REGION Network 4: alarmy
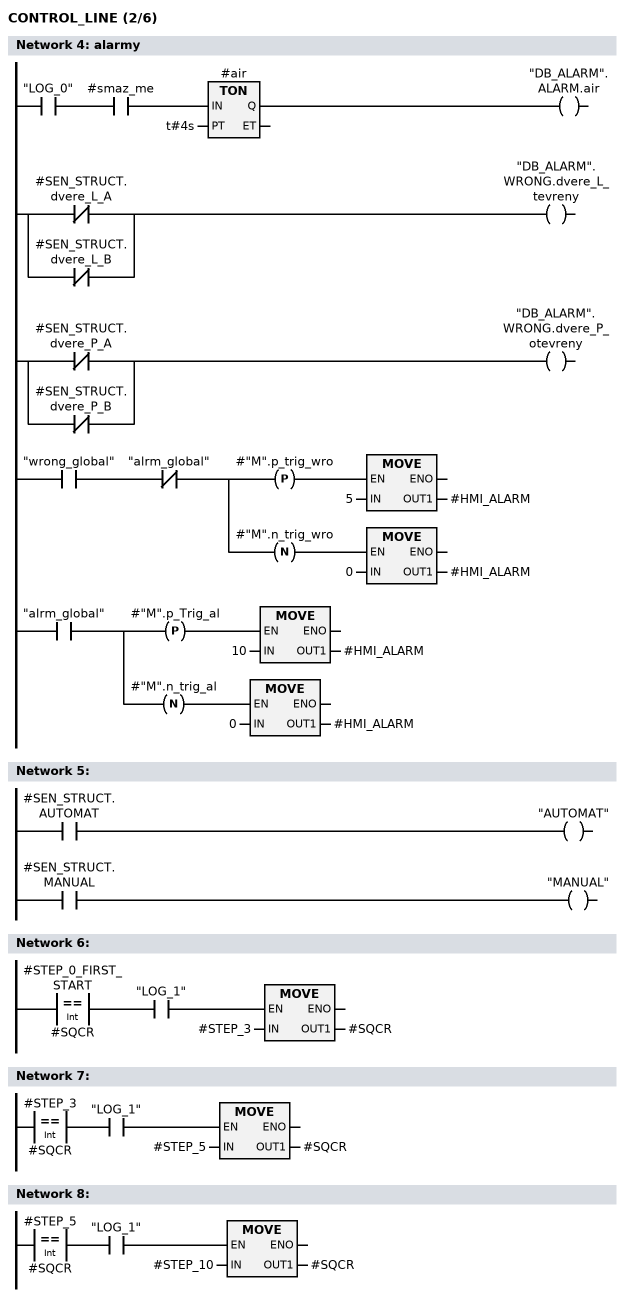
   #air(IN := "LOG_0" AND #smaz_me, PT := t#4s);   // TON
   "DB_ALARM".ALARM.air := #air.Q;
   "DB_ALARM".WRONG.dvere_L_tevreny := NOT #SEN_STRUCT.dvere_L_A OR NOT #SEN_STRUCT.dvere_L_B;
   "DB_ALARM".WRONG.dvere_P_otevreny := NOT #SEN_STRUCT.dvere_P_A OR NOT #SEN_STRUCT.dvere_P_B;
   #_w1 := "wrong_global" AND NOT "alrm_global";
   #_w2 := #_w1 AND NOT #"M".p_trig_wro;   // rising edge
   #"M".p_trig_wro := #_w1;
   IF #_w2 THEN #HMI_ALARM := 5; END_IF;
   #_w3 := NOT #_w1 AND #"M".n_trig_wro;   // falling edge
   #"M".n_trig_wro := #_w1;
   IF #_w3 THEN #HMI_ALARM := 0; END_IF;
   #_w4 := "alrm_global" AND NOT #"M".p_Trig_al;   // rising edge
   #"M".p_Trig_al := "alrm_global";
   IF #_w4 THEN #HMI_ALARM := 10; END_IF;
   #_w5 := NOT "alrm_global" AND #"M".n_trig_al;   // falling edge
   #"M".n_trig_al := "alrm_global";
   IF #_w5 THEN #HMI_ALARM := 0; END_IF;
END_REGION

REGION Network 5
   RUNG wire#powerrail
      Contact( #SEN_STRUCT.AUTOMAT )
      Coil( "AUTOMAT" )
   END_RUNG
   RUNG wire#powerrail
      Contact( #SEN_STRUCT.MANUAL )
      Coil( "MANUAL" )
   END_RUNG
   // the same network as SCL:
   "AUTOMAT" := #SEN_STRUCT.AUTOMAT;
   "MANUAL" := #SEN_STRUCT.MANUAL;
END_REGION

REGION Network 6
   RUNG wire#powerrail
      { S7_Templates := "SrcType := Int" } EQ_Contact(in1 := #STEP_0_FIRST_START, in2 := #SQCR)
      Contact( "LOG_1" )
      Move(in := #STEP_3, out1 => #SQCR)
   END_RUNG
   // the same network as SCL:
   IF (#STEP_0_FIRST_START = #SQCR) AND "LOG_1" THEN #SQCR := #STEP_3; END_IF;
END_REGION

REGION Network 7
   RUNG wire#powerrail
      { S7_Templates := "SrcType := Int" } EQ_Contact(in1 := #STEP_3, in2 := #SQCR)
      Contact( "LOG_1" )
      Move(in := #STEP_5, out1 => #SQCR)
   END_RUNG
   // the same network as SCL:
   IF (#STEP_3 = #SQCR) AND "LOG_1" THEN #SQCR := #STEP_5; END_IF;
END_REGION

REGION Network 8
   RUNG wire#powerrail
      { S7_Templates := "SrcType := Int" } EQ_Contact(in1 := #STEP_5, in2 := #SQCR)
      Contact( "LOG_1" )
      Move(in := #STEP_10, out1 => #SQCR)
   END_RUNG
   // the same network as SCL:
   IF (#STEP_5 = #SQCR) AND "LOG_1" THEN #SQCR := #STEP_10; END_IF;
END_REGION

REGION Network 9
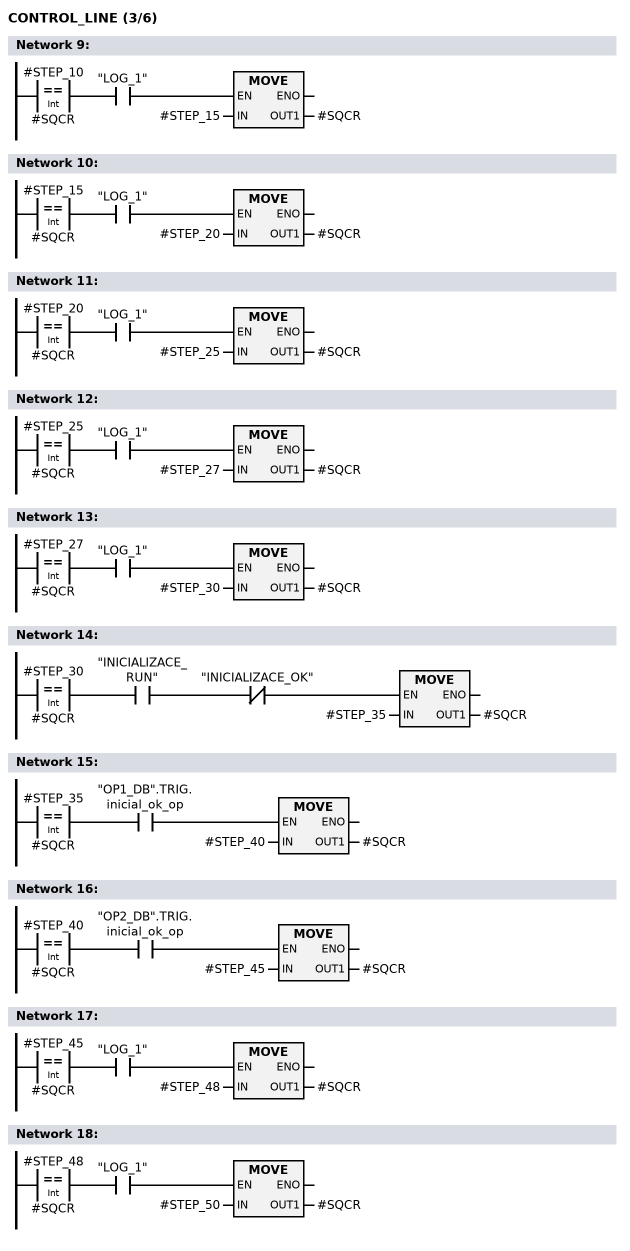
   RUNG wire#powerrail
      { S7_Templates := "SrcType := Int" } EQ_Contact(in1 := #STEP_10, in2 := #SQCR)
      Contact( "LOG_1" )
      Move(in := #STEP_15, out1 => #SQCR)
   END_RUNG
   // the same network as SCL:
   IF (#STEP_10 = #SQCR) AND "LOG_1" THEN #SQCR := #STEP_15; END_IF;
END_REGION

REGION Network 10
   RUNG wire#powerrail
      { S7_Templates := "SrcType := Int" } EQ_Contact(in1 := #STEP_15, in2 := #SQCR)
      Contact( "LOG_1" )
      Move(in := #STEP_20, out1 => #SQCR)
   END_RUNG
   // the same network as SCL:
   IF (#STEP_15 = #SQCR) AND "LOG_1" THEN #SQCR := #STEP_20; END_IF;
END_REGION

REGION Network 11
   RUNG wire#powerrail
      { S7_Templates := "SrcType := Int" } EQ_Contact(in1 := #STEP_20, in2 := #SQCR)
      Contact( "LOG_1" )
      Move(in := #STEP_25, out1 => #SQCR)
   END_RUNG
   // the same network as SCL:
   IF (#STEP_20 = #SQCR) AND "LOG_1" THEN #SQCR := #STEP_25; END_IF;
END_REGION

REGION Network 12
   RUNG wire#powerrail
      { S7_Templates := "SrcType := Int" } EQ_Contact(in1 := #STEP_25, in2 := #SQCR)
      Contact( "LOG_1" )
      Move(in := #STEP_27, out1 => #SQCR)
   END_RUNG
   // the same network as SCL:
   IF (#STEP_25 = #SQCR) AND "LOG_1" THEN #SQCR := #STEP_27; END_IF;
END_REGION

REGION Network 13
   RUNG wire#powerrail
      { S7_Templates := "SrcType := Int" } EQ_Contact(in1 := #STEP_27, in2 := #SQCR)
      Contact( "LOG_1" )
      Move(in := #STEP_30, out1 => #SQCR)
   END_RUNG
   // the same network as SCL:
   IF (#STEP_27 = #SQCR) AND "LOG_1" THEN #SQCR := #STEP_30; END_IF;
END_REGION

REGION Network 14
   RUNG wire#powerrail
      { S7_Templates := "SrcType := Int" } EQ_Contact(in1 := #STEP_30, in2 := #SQCR)
      Contact( "INICIALIZACE_RUN" )
      I_Contact( "INICIALIZACE_OK" )
      Move(in := #STEP_35, out1 => #SQCR)
   END_RUNG
   // the same network as SCL:
   IF (#STEP_30 = #SQCR) AND "INICIALIZACE_RUN" AND NOT "INICIALIZACE_OK" THEN #SQCR := #STEP_35; END_IF;
END_REGION

REGION Network 15
   RUNG wire#powerrail
      { S7_Templates := "SrcType := Int" } EQ_Contact(in1 := #STEP_35, in2 := #SQCR)
      Contact( "OP1_DB".TRIG.inicial_ok_op )
      Move(in := #STEP_40, out1 => #SQCR)
   END_RUNG
   // the same network as SCL:
   IF (#STEP_35 = #SQCR) AND "OP1_DB".TRIG.inicial_ok_op THEN #SQCR := #STEP_40; END_IF;
END_REGION

REGION Network 16
   RUNG wire#powerrail
      { S7_Templates := "SrcType := Int" } EQ_Contact(in1 := #STEP_40, in2 := #SQCR)
      Contact( "OP2_DB".TRIG.inicial_ok_op )
      Move(in := #STEP_45, out1 => #SQCR)
   END_RUNG
   // the same network as SCL:
   IF (#STEP_40 = #SQCR) AND "OP2_DB".TRIG.inicial_ok_op THEN #SQCR := #STEP_45; END_IF;
END_REGION

REGION Network 17
   RUNG wire#powerrail
      { S7_Templates := "SrcType := Int" } EQ_Contact(in1 := #STEP_45, in2 := #SQCR)
      Contact( "LOG_1" )
      Move(in := #STEP_48, out1 => #SQCR)
   END_RUNG
   // the same network as SCL:
   IF (#STEP_45 = #SQCR) AND "LOG_1" THEN #SQCR := #STEP_48; END_IF;
END_REGION

REGION Network 18
   RUNG wire#powerrail
      { S7_Templates := "SrcType := Int" } EQ_Contact(in1 := #STEP_48, in2 := #SQCR)
      Contact( "LOG_1" )
      Move(in := #STEP_50, out1 => #SQCR)
   END_RUNG
   // the same network as SCL:
   IF (#STEP_48 = #SQCR) AND "LOG_1" THEN #SQCR := #STEP_50; END_IF;
END_REGION

REGION Network 19
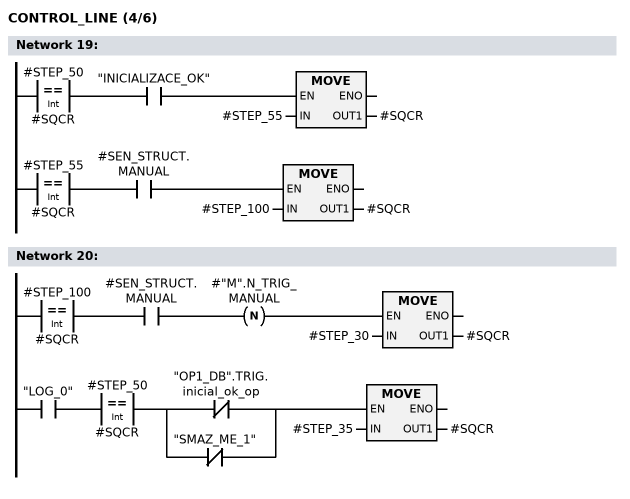
   RUNG wire#powerrail
      { S7_Templates := "SrcType := Int" } EQ_Contact(in1 := #STEP_50, in2 := #SQCR)
      Contact( "INICIALIZACE_OK" )
      Move(in := #STEP_55, out1 => #SQCR)
   END_RUNG
   RUNG wire#powerrail
      { S7_Templates := "SrcType := Int" } EQ_Contact(in1 := #STEP_55, in2 := #SQCR)
      Contact( #SEN_STRUCT.MANUAL )
      Move(in := #STEP_100, out1 => #SQCR)
   END_RUNG
   // the same network as SCL:
   IF (#STEP_50 = #SQCR) AND "INICIALIZACE_OK" THEN #SQCR := #STEP_55; END_IF;
   IF (#STEP_55 = #SQCR) AND #SEN_STRUCT.MANUAL THEN #SQCR := #STEP_100; END_IF;
END_REGION

REGION Network 20
   RUNG wire#powerrail
      { S7_Templates := "SrcType := Int" } EQ_Contact(in1 := #STEP_100, in2 := #SQCR)
      Contact( #SEN_STRUCT.MANUAL )
      N_Trig( #"M".N_TRIG_MANUAL )
      Move(in := #STEP_30, out1 => #SQCR)
   END_RUNG
   RUNG wire#powerrail
      Contact( "LOG_0" )
      { S7_Templates := "SrcType := Int" } EQ_Contact(in1 := #STEP_50, in2 := #SQCR)
      wire#w1
      I_Contact( "OP1_DB".TRIG.inicial_ok_op )
      wire#w2
      Move(in := #STEP_35, out1 => #SQCR)
   END_RUNG
   RUNG wire#w1
      I_Contact( "SMAZ_ME_1" )
   END_RUNG wire#w2
   // the same network as SCL:
   #_w1 := (#STEP_100 = #SQCR) AND #SEN_STRUCT.MANUAL;
   #_w2 := NOT #_w1 AND #"M".N_TRIG_MANUAL;   // falling edge
   #"M".N_TRIG_MANUAL := #_w1;
   IF #_w2 THEN #SQCR := #STEP_30; END_IF;
   IF "LOG_0" AND (#STEP_50 = #SQCR) AND (NOT "OP1_DB".TRIG.inicial_ok_op OR NOT "SMAZ_ME_1") THEN
       #SQCR := #STEP_35;
   END_IF;
END_REGION

REGION Network 21: LEDKY
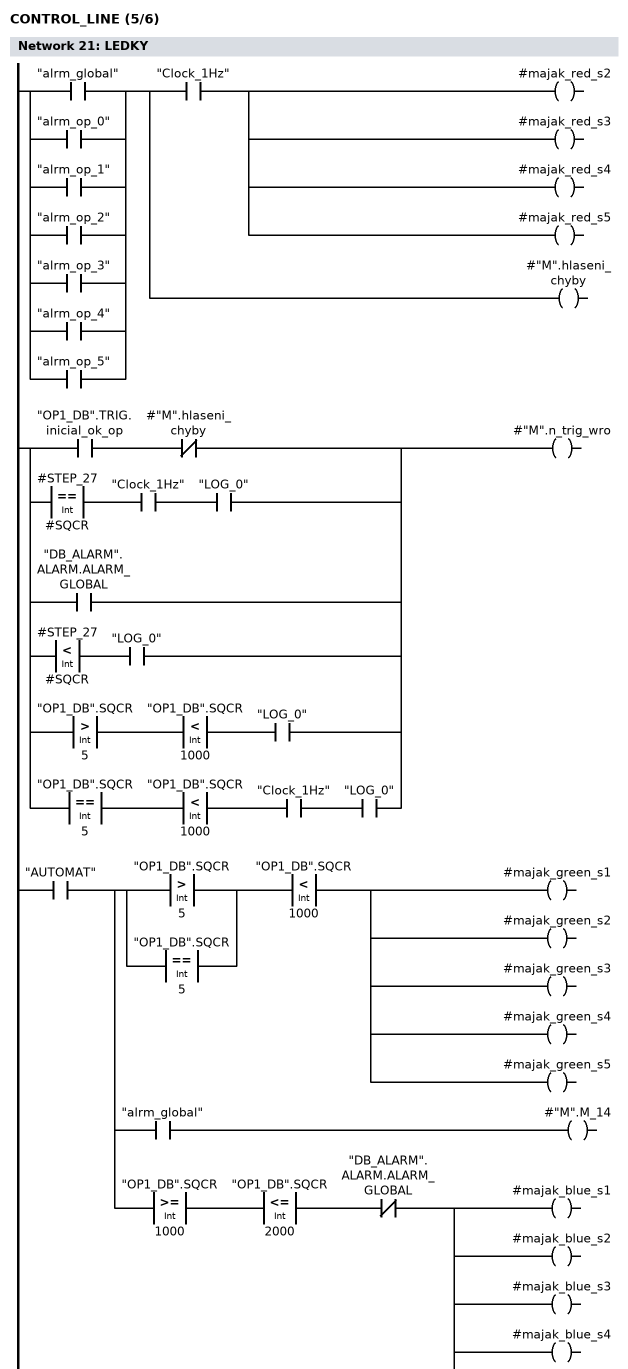
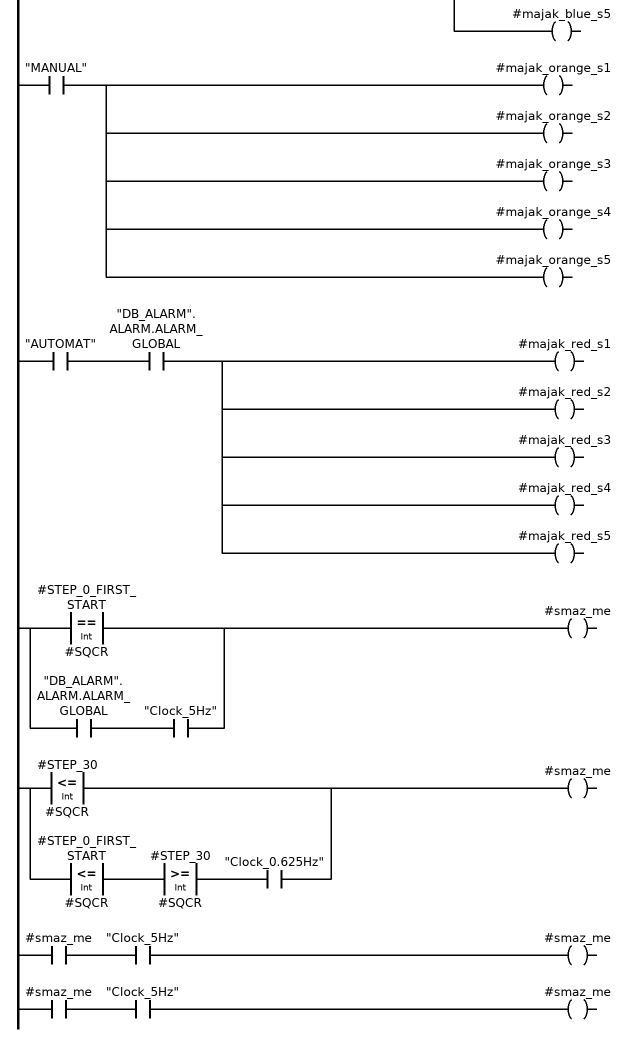
   RUNG wire#powerrail
      Contact( "alrm_global" )
      wire#w1
      Contact( "Clock_1Hz" )
      wire#w2
      Coil( #majak_red_s2 )
   END_RUNG
   RUNG wire#powerrail
      Contact( "alrm_op_0" )
   END_RUNG wire#w1
   RUNG wire#powerrail
      Contact( "alrm_op_1" )
   END_RUNG wire#w1
   RUNG wire#powerrail
      Contact( "alrm_op_2" )
   END_RUNG wire#w1
   RUNG wire#powerrail
      Contact( "alrm_op_3" )
   END_RUNG wire#w1
   RUNG wire#powerrail
      Contact( "alrm_op_4" )
   END_RUNG wire#w1
   RUNG wire#powerrail
      Contact( "alrm_op_5" )
   END_RUNG wire#w1
   RUNG wire#w2
      Coil( #majak_red_s3 )
   END_RUNG
   RUNG wire#w2
      Coil( #majak_red_s4 )
   END_RUNG
   RUNG wire#w2
      Coil( #majak_red_s5 )
   END_RUNG
   RUNG wire#w1
      Coil( #"M".hlaseni_chyby )
   END_RUNG
   RUNG wire#powerrail
      Contact( "OP1_DB".TRIG.inicial_ok_op )
      I_Contact( #"M".hlaseni_chyby )
      wire#w3
      Coil( #"M".n_trig_wro )
   END_RUNG
   RUNG wire#powerrail
      { S7_Templates := "SrcType := Int" } EQ_Contact(in1 := #STEP_27, in2 := #SQCR)
      Contact( "Clock_1Hz" )
      Contact( "LOG_0" )
   END_RUNG wire#w3
   RUNG wire#powerrail
      Contact( "DB_ALARM".ALARM.ALARM_GLOBAL )
   END_RUNG wire#w3
   RUNG wire#powerrail
      { S7_Templates := "SrcType := Int" } LT_Contact(in1 := #STEP_27, in2 := #SQCR)
      Contact( "LOG_0" )
   END_RUNG wire#w3
   RUNG wire#powerrail
      { S7_Templates := "SrcType := Int" } GT_Contact(in1 := "OP1_DB".SQCR, in2 := 5)
      { S7_Templates := "SrcType := Int" } LT_Contact(in1 := "OP1_DB".SQCR, in2 := 1000)
      Contact( "LOG_0" )
   END_RUNG wire#w3
   RUNG wire#powerrail
      { S7_Templates := "SrcType := Int" } EQ_Contact(in1 := "OP1_DB".SQCR, in2 := 5)
      { S7_Templates := "SrcType := Int" } LT_Contact(in1 := "OP1_DB".SQCR, in2 := 1000)
      Contact( "Clock_1Hz" )
      Contact( "LOG_0" )
   END_RUNG wire#w3
   RUNG wire#powerrail
      Contact( "AUTOMAT" )
      wire#w4
      { S7_Templates := "SrcType := Int" } GT_Contact(in1 := "OP1_DB".SQCR, in2 := 5)
      wire#w5
      { S7_Templates := "SrcType := Int" } LT_Contact(in1 := "OP1_DB".SQCR, in2 := 1000)
      wire#w6
      Coil( #majak_green_s1 )
   END_RUNG
   RUNG wire#w4
      { S7_Templates := "SrcType := Int" } EQ_Contact(in1 := "OP1_DB".SQCR, in2 := 5)
   END_RUNG wire#w5
   RUNG wire#w6
      Coil( #majak_green_s2 )
   END_RUNG
   RUNG wire#w6
      Coil( #majak_green_s3 )
   END_RUNG
   RUNG wire#w6
      Coil( #majak_green_s4 )
   END_RUNG
   RUNG wire#w6
      Coil( #majak_green_s5 )
   END_RUNG
   RUNG wire#w4
      Contact( "alrm_global" )
      Coil( #"M".M_14 )
   END_RUNG
   RUNG wire#w4
      { S7_Templates := "SrcType := Int" } GE_Contact(in1 := "OP1_DB".SQCR, in2 := 1000)
      { S7_Templates := "SrcType := Int" } LE_Contact(in1 := "OP1_DB".SQCR, in2 := 2000)
      I_Contact( "DB_ALARM".ALARM.ALARM_GLOBAL )
      wire#w7
      Coil( #majak_blue_s1 )
   END_RUNG
   RUNG wire#w7
      Coil( #majak_blue_s2 )
   END_RUNG
   RUNG wire#w7
      Coil( #majak_blue_s3 )
   END_RUNG
   RUNG wire#w7
      Coil( #majak_blue_s4 )
   END_RUNG
   RUNG wire#w7
      Coil( #majak_blue_s5 )
   END_RUNG
   RUNG wire#powerrail
      Contact( "MANUAL" )
      wire#w8
      Coil( #majak_orange_s1 )
   END_RUNG
   RUNG wire#w8
      Coil( #majak_orange_s2 )
   END_RUNG
   RUNG wire#w8
      Coil( #majak_orange_s3 )
   END_RUNG
   RUNG wire#w8
      Coil( #majak_orange_s4 )
   END_RUNG
   RUNG wire#w8
      Coil( #majak_orange_s5 )
   END_RUNG
   RUNG wire#powerrail
      Contact( "AUTOMAT" )
      Contact( "DB_ALARM".ALARM.ALARM_GLOBAL )
      wire#w9
      Coil( #majak_red_s1 )
   END_RUNG
   RUNG wire#w9
      Coil( #majak_red_s2 )
   END_RUNG
   RUNG wire#w9
      Coil( #majak_red_s3 )
   END_RUNG
   RUNG wire#w9
      Coil( #majak_red_s4 )
   END_RUNG
   RUNG wire#w9
      Coil( #majak_red_s5 )
   END_RUNG
   RUNG wire#powerrail
      { S7_Templates := "SrcType := Int" } EQ_Contact(in1 := #STEP_0_FIRST_START, in2 := #SQCR)
      wire#w10
      Coil( #smaz_me )
   END_RUNG
   RUNG wire#powerrail
      Contact( "DB_ALARM".ALARM.ALARM_GLOBAL )
      Contact( "Clock_5Hz" )
   END_RUNG wire#w10
   RUNG wire#powerrail
      { S7_Templates := "SrcType := Int" } LE_Contact(in1 := #STEP_30, in2 := #SQCR)
      wire#w11
      Coil( #smaz_me )
   END_RUNG
   RUNG wire#powerrail
      { S7_Templates := "SrcType := Int" } LE_Contact(in1 := #STEP_0_FIRST_START, in2 := #SQCR)
      { S7_Templates := "SrcType := Int" } GE_Contact(in1 := #STEP_30, in2 := #SQCR)
      Contact( "Clock_0.625Hz" )
   END_RUNG wire#w11
   RUNG wire#powerrail
      Contact( #smaz_me )
      Contact( "Clock_5Hz" )
      Coil( #smaz_me )
   END_RUNG
   RUNG wire#powerrail
      Contact( #smaz_me )
      Contact( "Clock_5Hz" )
      Coil( #smaz_me )
   END_RUNG
   // the same network as SCL:
   #_w1 := "alrm_global" OR "alrm_op_0" OR "alrm_op_1" OR "alrm_op_2" OR "alrm_op_3" OR "alrm_op_4" OR "alrm_op_5";
   #majak_red_s2 := #_w1 AND "Clock_1Hz";
   #majak_red_s3 := #majak_red_s2;
   #majak_red_s4 := #majak_red_s2;
   #majak_red_s5 := #majak_red_s2;
   #"M".hlaseni_chyby := #_w1;
   #"M".n_trig_wro := ("OP1_DB".TRIG.inicial_ok_op AND NOT #"M".hlaseni_chyby) OR ((#STEP_27 = #SQCR) AND "Clock_1Hz" AND "LOG_0") OR "DB_ALARM".ALARM.ALARM_GLOBAL OR ((#STEP_27 < #SQCR) AND "LOG_0") OR (("OP1_DB".SQCR > 5) AND ("OP1_DB".SQCR < 1000) AND "LOG_0") OR (("OP1_DB".SQCR = 5) AND ("OP1_DB".SQCR < 1000) AND "Clock_1Hz" AND "LOG_0");
   #majak_green_s1 := "AUTOMAT" AND (("OP1_DB".SQCR > 5) OR ("OP1_DB".SQCR = 5)) AND ("OP1_DB".SQCR < 1000);
   #majak_green_s2 := #majak_green_s1;
   #majak_green_s3 := #majak_green_s1;
   #majak_green_s4 := #majak_green_s1;
   #majak_green_s5 := #majak_green_s1;
   #"M".M_14 := "AUTOMAT" AND "alrm_global";
   #majak_blue_s1 := "AUTOMAT" AND ("OP1_DB".SQCR >= 1000) AND ("OP1_DB".SQCR <= 2000) AND NOT "DB_ALARM".ALARM.ALARM_GLOBAL;
   #majak_blue_s2 := #majak_blue_s1;
   #majak_blue_s3 := #majak_blue_s1;
   #majak_blue_s4 := #majak_blue_s1;
   #majak_blue_s5 := #majak_blue_s1;
   #majak_orange_s1 := "MANUAL";
   #majak_orange_s2 := "MANUAL";
   #majak_orange_s3 := "MANUAL";
   #majak_orange_s4 := "MANUAL";
   #majak_orange_s5 := "MANUAL";
   #majak_red_s1 := "AUTOMAT" AND "DB_ALARM".ALARM.ALARM_GLOBAL;
   #majak_red_s2 := #majak_red_s1;
   #majak_red_s3 := #majak_red_s1;
   #majak_red_s4 := #majak_red_s1;
   #majak_red_s5 := #majak_red_s1;
   #smaz_me := (#STEP_0_FIRST_START = #SQCR) OR ("DB_ALARM".ALARM.ALARM_GLOBAL AND "Clock_5Hz");
   #smaz_me := (#STEP_30 <= #SQCR) OR ((#STEP_0_FIRST_START <= #SQCR) AND (#STEP_30 >= #SQCR) AND "Clock_0.625Hz");
   #smaz_me := #smaz_me AND "Clock_5Hz";
   #smaz_me := #smaz_me AND "Clock_5Hz";
END_REGION

REGION Network 22: TRIG EXTERNAL
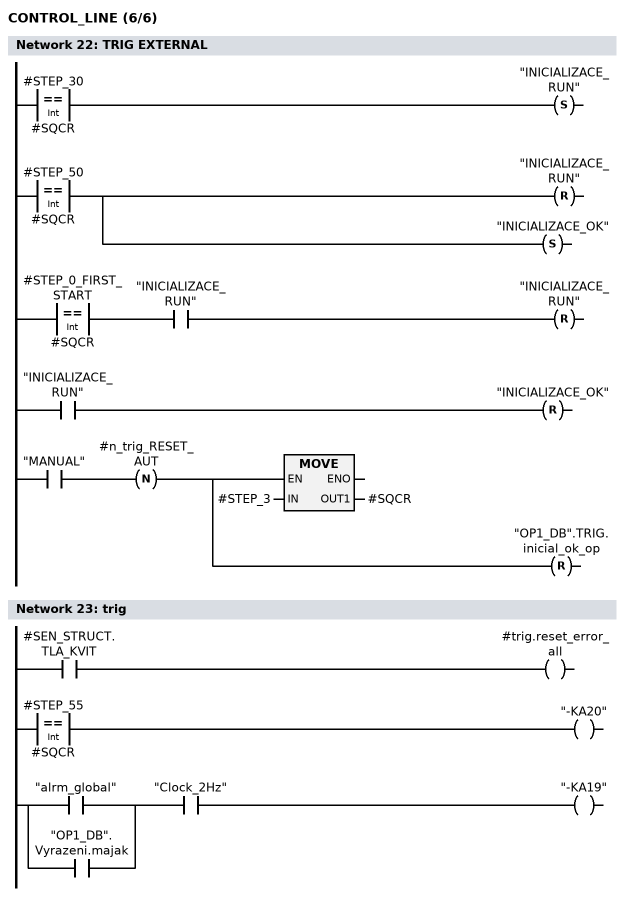
   RUNG wire#powerrail
      { S7_Templates := "SrcType := Int" } EQ_Contact(in1 := #STEP_30, in2 := #SQCR)
      S_Coil( "INICIALIZACE_RUN" )
   END_RUNG
   RUNG wire#powerrail
      { S7_Templates := "SrcType := Int" } EQ_Contact(in1 := #STEP_50, in2 := #SQCR)
      wire#w1
      R_Coil( "INICIALIZACE_RUN" )
   END_RUNG
   RUNG wire#w1
      S_Coil( "INICIALIZACE_OK" )
   END_RUNG
   RUNG wire#powerrail
      { S7_Templates := "SrcType := Int" } EQ_Contact(in1 := #STEP_0_FIRST_START, in2 := #SQCR)
      Contact( "INICIALIZACE_RUN" )
      R_Coil( "INICIALIZACE_RUN" )
   END_RUNG
   RUNG wire#powerrail
      Contact( "INICIALIZACE_RUN" )
      R_Coil( "INICIALIZACE_OK" )
   END_RUNG
   RUNG wire#powerrail
      Contact( "MANUAL" )
      N_Trig( #n_trig_RESET_AUT )
      wire#w2
      Move(in := #STEP_3, out1 => #SQCR)
   END_RUNG
   RUNG wire#w2
      R_Coil( "OP1_DB".TRIG.inicial_ok_op )
   END_RUNG
   // the same network as SCL:
   IF #STEP_30 = #SQCR THEN "INICIALIZACE_RUN" := TRUE; END_IF;
   IF #STEP_50 = #SQCR THEN
       "INICIALIZACE_RUN" := FALSE;
       "INICIALIZACE_OK" := TRUE;
   END_IF;
   IF (#STEP_0_FIRST_START = #SQCR) AND "INICIALIZACE_RUN" THEN "INICIALIZACE_RUN" := FALSE; END_IF;
   IF "INICIALIZACE_RUN" THEN "INICIALIZACE_OK" := FALSE; END_IF;
   #_w1 := NOT "MANUAL" AND #n_trig_RESET_AUT;   // falling edge
   #n_trig_RESET_AUT := "MANUAL";
   IF #_w1 THEN
       #SQCR := #STEP_3;
       "OP1_DB".TRIG.inicial_ok_op := FALSE;
   END_IF;
END_REGION

REGION Network 23: trig
   RUNG wire#powerrail
      Contact( #SEN_STRUCT.TLA_KVIT )
      Coil( #trig.reset_error_all )
   END_RUNG
   RUNG wire#powerrail
      { S7_Templates := "SrcType := Int" } EQ_Contact(in1 := #STEP_55, in2 := #SQCR)
      Coil( "-KA20" )
   END_RUNG
   RUNG wire#powerrail
      Contact( "alrm_global" )
      wire#w1
      Contact( "Clock_2Hz" )
      Coil( "-KA19" )
   END_RUNG
   RUNG wire#powerrail
      Contact( "OP1_DB".Vyrazeni.majak )
   END_RUNG wire#w1
   // the same network as SCL:
   #trig.reset_error_all := #SEN_STRUCT.TLA_KVIT;
   "-KA20" := #STEP_55 = #SQCR;
   "-KA19" := ("alrm_global" OR "OP1_DB".Vyrazeni.majak) AND "Clock_2Hz";
END_REGION
END_FUNCTION_BLOCK

(* ===== HMI "HMI_RT_1" =====
system functions are stored by id; their names below are inferred from use
connection "HMI_Connection_1": ETHERNET, SMART_S7_1200_OMS

HMI tags "Default tag table"
   "OP1_DB.Kamera.kontrola_tridirny" : Bool = PLC OP1_DB.Kamera.kontrola_tridirny, 1 s
   "alrm_global" : Bool = PLC alrm_global AT %M3.2, 1 s
   "AUT_MAN_HMI" : Bool = PLC AUT_MAN_HMI AT %M4.7, 1 s
   "CONTROL_LINE_DB_SQCR" : Int = PLC CONTROL_LINE_DB.SQCR, 1 s
   "DB_HMI_recype_recipe_Zprava" : Int = PLC DB_HMI_recype.recipe.Zprava, 1 s
   "DB_HMI_recype_recipe_PRG_CAM_etiketa" : Int = PLC DB_HMI_recype.recipe.PRG_CAM_etiketa, 1 s
   "DB_HMI_recype_recipe_PRG_CAM_folie" : Int = PLC DB_HMI_recype.recipe.PRG_CAM_folie, 1 s
   "DB_HMI_recype_recipe_vyrazovac_on_off" : Bool = PLC DB_HMI_recype.recipe.vyrazovac_on_off, 1 s
   "DB_HMI_recype_recipe_variabilni_pole_on_off" : Bool = PLC DB_HMI_recype.recipe.variabilni_pole_on_off, 1 s
   "DB_HMI_recype_fronta{1}_prenaseny_text" : String[100] = PLC DB_HMI_recype.fronta[1].prenaseny_text, 1 s
   "DB_HMI_recype_fronta{1}_balik_den" : Int = PLC DB_HMI_recype.fronta[1].balik_den, 1 s
   "DB_HMI_recype_fronta{1}_vyrazeni" : Bool = PLC DB_HMI_recype.fronta[1].vyrazeni, 1 s
   "DB_HMI_recype_fronta{2}_prenaseny_text" : String[100] = PLC DB_HMI_recype.fronta[2].prenaseny_text, 1 s
   "DB_HMI_recype_fronta{2}_balik_den" : Int = PLC DB_HMI_recype.fronta[2].balik_den, 1 s
   "DB_HMI_recype_fronta{2}_vyrazeni" : Bool = PLC DB_HMI_recype.fronta[2].vyrazeni, 1 s
   "DB_HMI_recype_fronta{3}_prenaseny_text" : String[100] = PLC DB_HMI_recype.fronta[3].prenaseny_text, 1 s
   "DB_HMI_recype_fronta{3}_balik_den" : Int = PLC DB_HMI_recype.fronta[3].balik_den, 1 s
   "DB_HMI_recype_fronta{3}_vyrazeni" : Bool = PLC DB_HMI_recype.fronta[3].vyrazeni, 1 s
   "DB_HMI_recype_fronta{4}_prenaseny_text" : String[100] = PLC DB_HMI_recype.fronta[4].prenaseny_text, 1 s
   "DB_HMI_recype_fronta{4}_balik_den" : Int = PLC DB_HMI_recype.fronta[4].balik_den, 1 s
   "DB_HMI_recype_fronta{4}_vyrazeni" : Bool = PLC DB_HMI_recype.fronta[4].vyrazeni, 1 s
   "DB_HMI_recype_fronta{5}_prenaseny_text" : String[100] = PLC DB_HMI_recype.fronta[5].prenaseny_text, 1 s
   "DB_HMI_recype_fronta{5}_balik_den" : Int = PLC DB_HMI_recype.fronta[5].balik_den, 1 s
   "DB_HMI_recype_fronta{5}_vyrazeni" : Bool = PLC DB_HMI_recype.fronta[5].vyrazeni, 1 s
   "DB_HMI_recype_obsazenost_fronty" : Int = PLC DB_HMI_recype.obsazenost_fronty, 1 s
   "OP1_DB_SENSORS_prechod_1" : Bool = PLC OP1_DB.SENSORS.prechod_1, 1 s
   "OP1_DB_SENSORS_kontrola" : Bool = PLC OP1_DB.SENSORS.kontrola, 1 s
   "OP1_DB_SENSORS_prechod_2" : Bool = PLC OP1_DB.SENSORS.prechod_2, 1 s
   "OP1_DB_SENSORS_Pozice_vyrazovace" : Bool = PLC OP1_DB.SENSORS.Pozice_vyrazovace, 1 s
   "OP1_DB_SENSORS_Pozice_pistu" : Bool = PLC OP1_DB.SENSORS.Pozice_pistu, 1 s
   "HSC_1" : DWord = PLC HSC_1 AT %ID1000, 1 s
   "OP1_DB_aktual_kusy" : Int = PLC OP1_DB.Kamera.balik_den, 1 s
   "OP2_DB_SQCR" : Int = PLC OP2_DB.SQCR AT %DB1.DBW658, 1 s
   "OP1_DB_HMI_hmi_5" : Bool = PLC OP1_DB.HMI.reset_fronty, 1 s
   "DB_HMI_recype_recipe_pole_string_1" : String[20] = PLC DB_HMI_recype.recipe.pole_string_1, 1 s
   "DB_HMI_recype_recipe_pole_string_2" : String[10] = PLC DB_HMI_recype.recipe.pole_string_2, 1 s
   "OP2_DB_TRIG_inicial_ok_op" : Bool = PLC OP2_DB.TRIG.inicial_ok_op AT %DB1.DBX662.0, 1 s
   "OP1_DB_SQCR" : Int = PLC OP1_DB.SQCR, 1 s
   "DB_HMI_recype_VZDALENOST_KAMERA_ETIKETA_POZADOVANA" : DInt = PLC DB_HMI_recype.VZDALENOST_KAMERA_ETIKETA_POZADOVANA, 1 s
   "DB_HMI_recype_VZDALENOST_KAMERY_FOLIE_POZADOVANA" : DInt = PLC DB_HMI_recype.VZDALENOST_KAMERY_FOLIE_POZADOVANA, 1 s
   "CONTROL_LINE_DB_HMI_ALARM" : Int = PLC CONTROL_LINE_DB.HMI_ALARM, 1 s
   "CONTROL_LINE_DB_SEN_STRUCT_dvere_L_A" : Bool = PLC CONTROL_LINE_DB.SEN_STRUCT.dvere_L_A, 1 s
   "CONTROL_LINE_DB_SEN_STRUCT_dvere_P_A" : Bool = PLC CONTROL_LINE_DB.SEN_STRUCT.dvere_P_A, 1 s
   "CONTROL_LINE_DB_SEN_STRUCT_dvere_L_B" : Bool = PLC CONTROL_LINE_DB.SEN_STRUCT.dvere_L_B, 1 s
   "CONTROL_LINE_DB_SEN_STRUCT_dvere_P_B" : Bool = PLC CONTROL_LINE_DB.SEN_STRUCT.dvere_P_B, 1 s
   "DB_HMI_recype_ODESLI_dATA" : Bool = PLC DB_HMI_recype.ODESLI_dATA, 100 ms
   "OK_Kusy_Den" : UInt, internal
   "NOK_Kusy_Den" : UInt, internal

HMI tags "alarmy"
   "DB_ALARM_OP1_M_0" : Int = PLC DB_ALARM.OP1.-Y7_KARUSEL AT %DB100.DBW44, 1 s
   "DB_ALARM_OP1_M_1" : Int = PLC DB_ALARM.OP1.-Y9_ZARAZKA AT %DB100.DBW46, 1 s
   "DB_ALARM_OP1_M_2" : Int = PLC DB_ALARM.OP1.M_2 AT %DB100.DBW48, 1 s
   "DB_ALARM_OP1_M_3" : Int = PLC DB_ALARM.OP1.M_3 AT %DB100.DBW50, 1 s
   "DB_ALARM_OP1_M_4" : Int = PLC DB_ALARM.OP1.M_4 AT %DB100.DBW52, 1 s
   "DB_ALARM_OP1_M_5" : Int = PLC DB_ALARM.OP1.M_5 AT %DB100.DBW54, 1 s
   "DB_ALARM_OP1_M_6" : Int = PLC DB_ALARM.OP1.M_6 AT %DB100.DBW56, 1 s
   "DB_ALARM_OP1_M_7" : Int = PLC DB_ALARM.OP1.M_7 AT %DB100.DBW58, 1 s
   "DB_ALARM_OP1_M_8" : Int = PLC DB_ALARM.OP1.M_8 AT %DB100.DBW60, 1 s
   "DB_ALARM_OP1_M_9" : Int = PLC DB_ALARM.OP1.M_9 AT %DB100.DBW62, 1 s
   "DB_ALARM_OP1_M_10" : Int = PLC DB_ALARM.OP1.M_10 AT %DB100.DBW64, 1 s
   "DB_ALARM_OP1_M_11" : Int = PLC DB_ALARM.OP1.M_11 AT %DB100.DBW66, 1 s
   "DB_ALARM_OP1_M_12" : Int = PLC DB_ALARM.OP1.M_12 AT %DB100.DBW68, 1 s
   "DB_ALARM_OP1_M_13" : Int = PLC DB_ALARM.OP1.M_13 AT %DB100.DBW70, 1 s
   "DB_ALARM_OP1_M_14" : Int = PLC DB_ALARM.OP1.M_14 AT %DB100.DBW72, 1 s
   "DB_ALARM_OP1_M_15" : Int = PLC DB_ALARM.OP1.M_15 AT %DB100.DBW74, 1 s
   "DB_ALARM_OP2_M_0" : Int = PLC DB_ALARM.OP2.A1 AT %DB100.DBW80, 1 s
   "DB_ALARM_OP2_M_1" : Int = PLC DB_ALARM.OP2.A2 AT %DB100.DBW82, 1 s
   "DB_ALARM_OP2_M_2" : Int = PLC DB_ALARM.OP2.A3 AT %DB100.DBW84, 1 s
   "DB_ALARM_OP2_M_3" : Int = PLC DB_ALARM.OP2.A4 AT %DB100.DBW86, 1 s
   "DB_ALARM_OP2_M_4" : Int = PLC DB_ALARM.OP2.A5 AT %DB100.DBW88, 1 s
   "DB_ALARM_OP2_M_5" : Int = PLC DB_ALARM.OP2.A6 AT %DB100.DBW90, 1 s
   "DB_ALARM_OP2_M_6" : Int = PLC DB_ALARM.OP2.A7 AT %DB100.DBW92, 1 s
   "DB_ALARM_OP2_M_7" : Int = PLC DB_ALARM.OP2.A8 AT %DB100.DBW94, 1 s
   "DB_ALARM_OP2_M_8" : Int = PLC DB_ALARM.OP2.M_8 AT %DB100.DBW96, 1 s
   "DB_ALARM_OP2_M_9" : Int = PLC DB_ALARM.OP2.M_9 AT %DB100.DBW98, 1 s
   "DB_ALARM_OP2_M_10" : Int = PLC DB_ALARM.OP2.M_10 AT %DB100.DBW100, 1 s
   "DB_ALARM_OP2_M_11" : Int = PLC DB_ALARM.OP2.M_11 AT %DB100.DBW102, 1 s
   "DB_ALARM_OP2_M_12" : Int = PLC DB_ALARM.OP2.M_12 AT %DB100.DBW104, 1 s
   "DB_ALARM_OP2_M_13" : Int = PLC DB_ALARM.OP2.M_13 AT %DB100.DBW106, 1 s
   "DB_ALARM_OP2_M_14" : Int = PLC DB_ALARM.OP2.M_14 AT %DB100.DBW108, 1 s
   "DB_ALARM_OP2_M_15" : Int = PLC DB_ALARM.OP2.M_15 AT %DB100.DBW110, 1 s
   "DB_ALARM_OP3_M_0" : Int = PLC DB_ALARM.OP3.B1 AT %DB100.DBW116, 1 s
   "DB_ALARM_OP3_M_1" : Int = PLC DB_ALARM.OP3.B2 AT %DB100.DBW118, 1 s
   "DB_ALARM_OP3_M_2" : Int = PLC DB_ALARM.OP3.B3 AT %DB100.DBW120, 1 s
   "DB_ALARM_OP3_M_3" : Int = PLC DB_ALARM.OP3.B4 AT %DB100.DBW122, 1 s
   "DB_ALARM_OP3_M_4" : Int = PLC DB_ALARM.OP3.B5 AT %DB100.DBW124, 1 s
   "DB_ALARM_OP3_M_5" : Int = PLC DB_ALARM.OP3.B6 AT %DB100.DBW126, 1 s
   "DB_ALARM_OP3_M_6" : Int = PLC DB_ALARM.OP3.B7 AT %DB100.DBW128, 1 s
   "DB_ALARM_OP3_M_7" : Int = PLC DB_ALARM.OP3.B8 AT %DB100.DBW130, 1 s
   "DB_ALARM_OP3_M_8" : Int = PLC DB_ALARM.OP3.M_8 AT %DB100.DBW132, 1 s
   "DB_ALARM_OP3_M_9" : Int = PLC DB_ALARM.OP3.M_9 AT %DB100.DBW134, 1 s
   "DB_ALARM_OP3_M_10" : Int = PLC DB_ALARM.OP3.M_10 AT %DB100.DBW136, 1 s
   "DB_ALARM_OP3_M_11" : Int = PLC DB_ALARM.OP3.M_11 AT %DB100.DBW138, 1 s
   "DB_ALARM_OP3_M_12" : Int = PLC DB_ALARM.OP3.M_12 AT %DB100.DBW140, 1 s
   "DB_ALARM_OP3_M_13" : Int = PLC DB_ALARM.OP3.M_13 AT %DB100.DBW142, 1 s
   "DB_ALARM_OP3_M_14" : Int = PLC DB_ALARM.OP3.M_14 AT %DB100.DBW144, 1 s
   "DB_ALARM_OP3_M_15" : Int = PLC DB_ALARM.OP3.M_15 AT %DB100.DBW146, 1 s
   "DB_ALARM_OP1_ALARM_dvere_1" : Bool = PLC DB_ALARM.OP1.ALARM.dvere_1 AT %DB100.DBX40.0, 1 s
   "DB_ALARM_OP1_ALARM_ALARM_1" : Bool = PLC DB_ALARM.OP1.ALARM.ALARM_1 AT %DB100.DBX40.1, 1 s
   "DB_ALARM_OP1_ALARM_ALARM_2" : Bool = PLC DB_ALARM.OP1.ALARM.ALARM_2 AT %DB100.DBX40.2, 1 s
   "DB_ALARM_OP1_ALARM_ALARM_3" : Bool = PLC DB_ALARM.OP1.ALARM.ALARM_3 AT %DB100.DBX40.3, 1 s
   "DB_ALARM_OP1_ALARM_ALARM_4" : Bool = PLC DB_ALARM.OP1.ALARM.ALARM_4 AT %DB100.DBX40.4, 1 s
   "DB_ALARM_OP1_ALARM_ALARM_5" : Bool = PLC DB_ALARM.OP1.ALARM.ALARM_5 AT %DB100.DBX40.5, 1 s
   "DB_ALARM_OP1_ALARM_ALARM_6" : Bool = PLC DB_ALARM.OP1.ALARM.ALARM_6 AT %DB100.DBX40.6, 1 s
   "DB_ALARM_OP1_ALARM_hladina_mimo_mez" : Bool = PLC DB_ALARM.OP1.ALARM.hladina_mimo_mez AT %DB100.DBX40.7, 1 s
   "DB_ALARM_OP1_ALARM_ALARM_8" : Bool = PLC DB_ALARM.OP1.ALARM.ALARM_8 AT %DB100.DBX41.0, 1 s
   "DB_ALARM_OP1_ALARM_ALARM_9" : Bool = PLC DB_ALARM.OP1.ALARM.ALARM_9 AT %DB100.DBX41.1, 1 s
   "DB_ALARM_OP1_ALARM_ALARM_10" : Bool = PLC DB_ALARM.OP1.ALARM.ALARM_10 AT %DB100.DBX41.2, 1 s
   "DB_ALARM_OP1_ALARM_ALARM_11" : Bool = PLC DB_ALARM.OP1.ALARM.ALARM_11 AT %DB100.DBX41.3, 1 s
   "DB_ALARM_OP1_ALARM_ALARM_12" : Bool = PLC DB_ALARM.OP1.ALARM.ALARM_12 AT %DB100.DBX41.4, 1 s
   "DB_ALARM_OP1_ALARM_ALARM_13" : Bool = PLC DB_ALARM.OP1.ALARM.ALARM_13 AT %DB100.DBX41.5, 1 s
   "DB_ALARM_OP1_ALARM_ALARM_14" : Bool = PLC DB_ALARM.OP1.ALARM.ALARM_14 AT %DB100.DBX41.6, 1 s
   "DB_ALARM_OP1_ALARM_ALARM_15" : Bool = PLC DB_ALARM.OP1.ALARM.ALARM_15 AT %DB100.DBX41.7, 1 s
   "DB_ALARM_OP2_ALARM_dvere_1" : Bool = PLC DB_ALARM.OP2.ALARM.dvere_1 AT %DB100.DBX76.0, 1 s
   "DB_ALARM_OP2_ALARM_dvere_2" : Bool = PLC DB_ALARM.OP2.ALARM.dvere_2 AT %DB100.DBX76.1, 1 s
   "DB_ALARM_OP2_ALARM_dvere_3" : Bool = PLC DB_ALARM.OP2.ALARM.dvere_3 AT %DB100.DBX76.2, 1 s
   "DB_ALARM_OP2_ALARM_dvere_4" : Bool = PLC DB_ALARM.OP2.ALARM.dvere_4 AT %DB100.DBX76.3, 1 s
   "DB_ALARM_OP2_ALARM_paprsek" : Bool = PLC DB_ALARM.OP2.ALARM.paprsek AT %DB100.DBX76.4, 1 s
   "DB_ALARM_OP2_ALARM_porucha_svarovani" : Bool = PLC DB_ALARM.OP2.ALARM.porucha_svarovani AT %DB100.DBX76.5, 1 s
   "DB_ALARM_OP2_ALARM_rop_alarm" : Bool = PLC DB_ALARM.OP2.ALARM.rop_alarm AT %DB100.DBX76.6, 1 s
   "DB_ALARM_OP2_ALARM_servo_power_error" : Bool = PLC DB_ALARM.OP2.ALARM.servo_power_error AT %DB100.DBX76.7, 1 s
   "DB_ALARM_OP2_ALARM_servo_jog_error" : Bool = PLC DB_ALARM.OP2.ALARM.servo_jog_error AT %DB100.DBX77.0, 1 s
   "DB_ALARM_OP2_ALARM_servo_homing" : Bool = PLC DB_ALARM.OP2.ALARM.servo_homing AT %DB100.DBX77.1, 1 s
   "DB_ALARM_OP2_ALARM_Cel_podel_porucha" : Bool = PLC DB_ALARM.OP2.ALARM.Cel_podel_porucha AT %DB100.DBX77.2, 1 s
   "DB_ALARM_OP2_ALARM_vysoka_tuzka" : Bool = PLC DB_ALARM.OP2.ALARM.vysoka_tuzka AT %DB100.DBX77.3, 1 s
   "DB_ALARM_OP2_ALARM_ALARM_12" : Bool = PLC DB_ALARM.OP2.ALARM.ALARM_12 AT %DB100.DBX77.4, 1 s
   "DB_ALARM_OP2_ALARM_ALARM_13" : Bool = PLC DB_ALARM.OP2.ALARM.ALARM_13 AT %DB100.DBX77.5, 1 s
   "DB_ALARM_OP2_ALARM_folie" : Bool = PLC DB_ALARM.OP2.ALARM.folie AT %DB100.DBX77.6, 1 s
   "DB_ALARM_OP2_ALARM_ALARM_15" : Bool = PLC DB_ALARM.OP2.ALARM.ALARM_15 AT %DB100.DBX77.7, 1 s
   "DB_ALARM_OP3_ALARM_ALARM_0" : Bool = PLC DB_ALARM.OP3.ALARM.ALARM_0 AT %DB100.DBX112.0, 1 s
   "DB_ALARM_OP3_ALARM_ALARM_1" : Bool = PLC DB_ALARM.OP3.ALARM.ALARM_1 AT %DB100.DBX112.1, 1 s
   "DB_ALARM_OP3_ALARM_ALARM_2" : Bool = PLC DB_ALARM.OP3.ALARM.ALARM_2 AT %DB100.DBX112.2, 1 s
   "DB_ALARM_OP3_ALARM_ALARM_3" : Bool = PLC DB_ALARM.OP3.ALARM.ALARM_3 AT %DB100.DBX112.3, 1 s
   "DB_ALARM_OP3_ALARM_ALARM_4" : Bool = PLC DB_ALARM.OP3.ALARM.ALARM_4 AT %DB100.DBX112.4, 1 s
   "DB_ALARM_OP3_ALARM_ALARM_5" : Bool = PLC DB_ALARM.OP3.ALARM.ALARM_5 AT %DB100.DBX112.5, 1 s
   "DB_ALARM_OP3_ALARM_ALARM_6" : Bool = PLC DB_ALARM.OP3.ALARM.ALARM_6 AT %DB100.DBX112.6, 1 s
   "DB_ALARM_OP3_ALARM_ALARM_7" : Bool = PLC DB_ALARM.OP3.ALARM.ALARM_7 AT %DB100.DBX112.7, 1 s
   "DB_ALARM_OP3_ALARM_ALARM_8" : Bool = PLC DB_ALARM.OP3.ALARM.ALARM_8 AT %DB100.DBX113.0, 1 s
   "DB_ALARM_OP3_ALARM_ALARM_9" : Bool = PLC DB_ALARM.OP3.ALARM.ALARM_9 AT %DB100.DBX113.1, 1 s
   "DB_ALARM_OP3_ALARM_ALARM_10" : Bool = PLC DB_ALARM.OP3.ALARM.ALARM_10 AT %DB100.DBX113.2, 1 s
   "DB_ALARM_OP3_ALARM_ALARM_11" : Bool = PLC DB_ALARM.OP3.ALARM.ALARM_11 AT %DB100.DBX113.3, 1 s
   "DB_ALARM_OP3_ALARM_ALARM_12" : Bool = PLC DB_ALARM.OP3.ALARM.ALARM_12 AT %DB100.DBX113.4, 1 s
   "DB_ALARM_OP3_ALARM_ALARM_13" : Bool = PLC DB_ALARM.OP3.ALARM.ALARM_13 AT %DB100.DBX113.5, 1 s
   "DB_ALARM_OP3_ALARM_ALARM_14" : Bool = PLC DB_ALARM.OP3.ALARM.ALARM_14 AT %DB100.DBX113.6, 1 s
   "DB_ALARM_OP3_ALARM_ALARM_15" : Bool = PLC DB_ALARM.OP3.ALARM.ALARM_15 AT %DB100.DBX113.7, 1 s
   "DB_ALARM_OP1_WRONG_WRONG_0" : Bool = PLC DB_ALARM.OP1.WRONG.WRONG_0 AT %DB100.DBX42.0, 1 s
   "DB_ALARM_OP1_WRONG_WRONG_1" : Bool = PLC DB_ALARM.OP1.WRONG.WRONG_1 AT %DB100.DBX42.1, 1 s
   "DB_ALARM_OP1_WRONG_WRONG_2" : Bool = PLC DB_ALARM.OP1.WRONG.WRONG_2 AT %DB100.DBX42.2, 1 s
   "DB_ALARM_OP1_WRONG_WRONG_3" : Bool = PLC DB_ALARM.OP1.WRONG.WRONG_3 AT %DB100.DBX42.3, 1 s
   "DB_ALARM_OP1_WRONG_WRONG_4" : Bool = PLC DB_ALARM.OP1.WRONG.WRONG_4 AT %DB100.DBX42.4, 1 s
   "DB_ALARM_OP1_WRONG_WRONG_5" : Bool = PLC DB_ALARM.OP1.WRONG.WRONG_5 AT %DB100.DBX42.5, 1 s
   "DB_ALARM_OP1_WRONG_WRONG_6" : Bool = PLC DB_ALARM.OP1.WRONG.WRONG_6 AT %DB100.DBX42.6, 1 s
   "DB_ALARM_OP1_WRONG_WRONG_7" : Bool = PLC DB_ALARM.OP1.WRONG.WRONG_7 AT %DB100.DBX42.7, 1 s
   "DB_ALARM_OP1_WRONG_WRONG_8" : Bool = PLC DB_ALARM.OP1.WRONG.WRONG_8 AT %DB100.DBX43.0, 1 s
   "DB_ALARM_OP1_WRONG_WRONG_9" : Bool = PLC DB_ALARM.OP1.WRONG.WRONG_9 AT %DB100.DBX43.1, 1 s
   "DB_ALARM_OP1_WRONG_WRONG_10" : Bool = PLC DB_ALARM.OP1.WRONG.WRONG_10 AT %DB100.DBX43.2, 1 s
   "DB_ALARM_OP1_WRONG_WRONG_11" : Bool = PLC DB_ALARM.OP1.WRONG.WRONG_11 AT %DB100.DBX43.3, 1 s
   "DB_ALARM_OP1_WRONG_WRONG_12" : Bool = PLC DB_ALARM.OP1.WRONG.WRONG_12 AT %DB100.DBX43.4, 1 s
   "DB_ALARM_OP1_WRONG_WRONG_13" : Bool = PLC DB_ALARM.OP1.WRONG.WRONG_13 AT %DB100.DBX43.5, 1 s
   "DB_ALARM_OP1_WRONG_WRONG_14" : Bool = PLC DB_ALARM.OP1.WRONG.WRONG_14 AT %DB100.DBX43.6, 1 s
   "DB_ALARM_OP1_WRONG_WRONG_15" : Bool = PLC DB_ALARM.OP1.WRONG.WRONG_15 AT %DB100.DBX43.7, 1 s
   "DB_ALARM_OP2_WRONG_WRONG_0" : Bool = PLC DB_ALARM.OP2.WRONG.WRONG_0 AT %DB100.DBX78.0, 1 s
   "DB_ALARM_OP2_WRONG_WRONG_1" : Bool = PLC DB_ALARM.OP2.WRONG.WRONG_1 AT %DB100.DBX78.1, 1 s
   "DB_ALARM_OP2_WRONG_WRONG_2" : Bool = PLC DB_ALARM.OP2.WRONG.WRONG_2 AT %DB100.DBX78.2, 1 s
   "DB_ALARM_OP2_WRONG_WRONG_3" : Bool = PLC DB_ALARM.OP2.WRONG.WRONG_3 AT %DB100.DBX78.3, 1 s
   "DB_ALARM_OP2_WRONG_WRONG_4" : Bool = PLC DB_ALARM.OP2.WRONG.WRONG_4 AT %DB100.DBX78.4, 1 s
   "DB_ALARM_OP2_WRONG_WRONG_5" : Bool = PLC DB_ALARM.OP2.WRONG.WRONG_5 AT %DB100.DBX78.5, 1 s
   "DB_ALARM_OP2_WRONG_WRONG_6" : Bool = PLC DB_ALARM.OP2.WRONG.WRONG_6 AT %DB100.DBX78.6, 1 s
   "DB_ALARM_OP2_WRONG_WRONG_7" : Bool = PLC DB_ALARM.OP2.WRONG.WRONG_7 AT %DB100.DBX78.7, 1 s
   "DB_ALARM_OP2_WRONG_WRONG_8" : Bool = PLC DB_ALARM.OP2.WRONG.WRONG_8 AT %DB100.DBX79.0, 1 s
   "DB_ALARM_OP2_WRONG_WRONG_9" : Bool = PLC DB_ALARM.OP2.WRONG.WRONG_9 AT %DB100.DBX79.1, 1 s
   "DB_ALARM_OP2_WRONG_WRONG_10" : Bool = PLC DB_ALARM.OP2.WRONG.WRONG_10 AT %DB100.DBX79.2, 1 s
   "DB_ALARM_OP2_WRONG_WRONG_11" : Bool = PLC DB_ALARM.OP2.WRONG.WRONG_11 AT %DB100.DBX79.3, 1 s
   "DB_ALARM_OP2_WRONG_WRONG_12" : Bool = PLC DB_ALARM.OP2.WRONG.WRONG_12 AT %DB100.DBX79.4, 1 s
   "DB_ALARM_OP2_WRONG_WRONG_13" : Bool = PLC DB_ALARM.OP2.WRONG.WRONG_13 AT %DB100.DBX79.5, 1 s
   "DB_ALARM_OP2_WRONG_WRONG_14" : Bool = PLC DB_ALARM.OP2.WRONG.WRONG_14 AT %DB100.DBX79.6, 1 s
   "DB_ALARM_OP2_WRONG_WRONG_15" : Bool = PLC DB_ALARM.OP2.WRONG.WRONG_15 AT %DB100.DBX79.7, 1 s
   "DB_ALARM_OP3_WRONG_WRONG_0" : Bool = PLC DB_ALARM.OP3.WRONG.WRONG_0 AT %DB100.DBX114.0, 1 s
   "DB_ALARM_OP3_WRONG_WRONG_1" : Bool = PLC DB_ALARM.OP3.WRONG.WRONG_1 AT %DB100.DBX114.1, 1 s
   "DB_ALARM_OP3_WRONG_WRONG_2" : Bool = PLC DB_ALARM.OP3.WRONG.WRONG_2 AT %DB100.DBX114.2, 1 s
   "DB_ALARM_OP3_WRONG_WRONG_3" : Bool = PLC DB_ALARM.OP3.WRONG.WRONG_3 AT %DB100.DBX114.3, 1 s
   "DB_ALARM_OP3_WRONG_WRONG_4" : Bool = PLC DB_ALARM.OP3.WRONG.WRONG_4 AT %DB100.DBX114.4, 1 s
   "DB_ALARM_OP3_WRONG_WRONG_5" : Bool = PLC DB_ALARM.OP3.WRONG.WRONG_5 AT %DB100.DBX114.5, 1 s
   "DB_ALARM_OP3_WRONG_WRONG_6" : Bool = PLC DB_ALARM.OP3.WRONG.WRONG_6 AT %DB100.DBX114.6, 1 s
   "DB_ALARM_OP3_WRONG_WRONG_7" : Bool = PLC DB_ALARM.OP3.WRONG.WRONG_7 AT %DB100.DBX114.7, 1 s
   "DB_ALARM_OP3_WRONG_WRONG_8" : Bool = PLC DB_ALARM.OP3.WRONG.WRONG_8 AT %DB100.DBX115.0, 1 s
   "DB_ALARM_OP3_WRONG_WRONG_9" : Bool = PLC DB_ALARM.OP3.WRONG.WRONG_9 AT %DB100.DBX115.1, 1 s
   "DB_ALARM_OP3_WRONG_WRONG_10" : Bool = PLC DB_ALARM.OP3.WRONG.WRONG_10 AT %DB100.DBX115.2, 1 s
   "DB_ALARM_OP3_WRONG_WRONG_11" : Bool = PLC DB_ALARM.OP3.WRONG.WRONG_11 AT %DB100.DBX115.3, 1 s
   "DB_ALARM_OP3_WRONG_WRONG_12" : Bool = PLC DB_ALARM.OP3.WRONG.WRONG_12 AT %DB100.DBX115.4, 1 s
   "DB_ALARM_OP3_WRONG_WRONG_13" : Bool = PLC DB_ALARM.OP3.WRONG.WRONG_13 AT %DB100.DBX115.5, 1 s
   "DB_ALARM_OP3_WRONG_WRONG_14" : Bool = PLC DB_ALARM.OP3.WRONG.WRONG_14 AT %DB100.DBX115.6, 1 s
   "DB_ALARM_OP3_WRONG_WRONG_15" : Bool = PLC DB_ALARM.OP3.WRONG.WRONG_15 AT %DB100.DBX115.7, 1 s
   "DB_ALARM_ALARM_ALARM_GLOBAL" : Bool = PLC DB_ALARM.ALARM.ALARM_GLOBAL AT %DB100.DBX0.0, 1 s
   "DB_ALARM_ALARM_HERMA_ERROR" : Bool = PLC DB_ALARM.ALARM.HERMA_ERROR AT %DB100.DBX0.1, 1 s
   "DB_ALARM_ALARM_ALARM_2" : Bool = PLC DB_ALARM.ALARM.ALARM_2 AT %DB100.DBX0.2, 1 s
   "DB_ALARM_ALARM_ALARM_3" : Bool = PLC DB_ALARM.ALARM.ALARM_3 AT %DB100.DBX0.3, 1 s
   "DB_ALARM_ALARM_ALARM_4" : Bool = PLC DB_ALARM.ALARM.ALARM_4 AT %DB100.DBX0.4, 1 s
   "DB_ALARM_ALARM_ALARM_5" : Bool = PLC DB_ALARM.ALARM.ALARM_5 AT %DB100.DBX0.5, 1 s
   "DB_ALARM_ALARM_air" : Bool = PLC DB_ALARM.ALARM.air AT %DB100.DBX0.6, 1 s
   "DB_ALARM_ALARM_ALARM_7" : Bool = PLC DB_ALARM.ALARM.ALARM_7 AT %DB100.DBX0.7, 1 s
   "DB_ALARM_ALARM_ALARM_8" : Bool = PLC DB_ALARM.ALARM.ALARM_8 AT %DB100.DBX1.0, 1 s
   "DB_ALARM_ALARM_ALARM_9" : Bool = PLC DB_ALARM.ALARM.ALARM_9 AT %DB100.DBX1.1, 1 s
   "DB_ALARM_ALARM_ALARM_10" : Bool = PLC DB_ALARM.ALARM.ALARM_10 AT %DB100.DBX1.2, 1 s
   "DB_ALARM_ALARM_ALARM_11" : Bool = PLC DB_ALARM.ALARM.ALARM_11 AT %DB100.DBX1.3, 1 s
   "DB_ALARM_ALARM_ALARM_12" : Bool = PLC DB_ALARM.ALARM.ALARM_12 AT %DB100.DBX1.4, 1 s
   "DB_ALARM_ALARM_ALARM_13" : Bool = PLC DB_ALARM.ALARM.ALARM_13 AT %DB100.DBX1.5, 1 s
   "DB_ALARM_ALARM_ALARM_14" : Bool = PLC DB_ALARM.ALARM.ALARM_14 AT %DB100.DBX1.6, 1 s
   "DB_ALARM_ALARM_vypadek_safety_karty" : Bool = PLC DB_ALARM.ALARM.vypadek_safety_karty AT %DB100.DBX1.7, 1 s
   "DB_ALARM_WRONG_NENI_INICIALIZACE" : Bool = PLC DB_ALARM.WRONG.NENI_INICIALIZACE AT %DB100.DBX2.0, 1 s
   "DB_ALARM_WRONG_WRONG_global" : Bool = PLC DB_ALARM.WRONG.WRONG_global AT %DB100.DBX2.1, 1 s
   "DB_ALARM_WRONG_WRONG_2" : Bool = PLC DB_ALARM.WRONG.dvere_L_tevreny AT %DB100.DBX2.2, 1 s
   "DB_ALARM_WRONG_WRONG_3" : Bool = PLC DB_ALARM.WRONG.dvere_P_otevreny AT %DB100.DBX2.3, 1 s
   "DB_ALARM_WRONG_WRONG_4" : Bool = PLC DB_ALARM.WRONG.WRONG_4 AT %DB100.DBX2.4, 1 s
   "DB_ALARM_WRONG_WRONG_5" : Bool = PLC DB_ALARM.WRONG.WRONG_5 AT %DB100.DBX2.5, 1 s
   "DB_ALARM_WRONG_WRONG_6" : Bool = PLC DB_ALARM.WRONG.WRONG_6 AT %DB100.DBX2.6, 1 s
   "DB_ALARM_WRONG_WRONG_7" : Bool = PLC DB_ALARM.WRONG.WRONG_7 AT %DB100.DBX2.7, 1 s
   "DB_ALARM_WRONG_WRONG_8" : Bool = PLC DB_ALARM.WRONG.WRONG_8 AT %DB100.DBX3.0, 1 s
   "DB_ALARM_WRONG_WRONG_9" : Bool = PLC DB_ALARM.WRONG.WRONG_9 AT %DB100.DBX3.1, 1 s
   "DB_ALARM_WRONG_WRONG_10" : Bool = PLC DB_ALARM.WRONG.WRONG_10 AT %DB100.DBX3.2, 1 s
   "DB_ALARM_WRONG_WRONG_11" : Bool = PLC DB_ALARM.WRONG.WRONG_11 AT %DB100.DBX3.3, 1 s
   "DB_ALARM_WRONG_WRONG_12" : Bool = PLC DB_ALARM.WRONG.WRONG_12 AT %DB100.DBX3.4, 1 s
   "DB_ALARM_WRONG_WRONG_13" : Bool = PLC DB_ALARM.WRONG.WRONG_13 AT %DB100.DBX3.5, 1 s
   "DB_ALARM_WRONG_rop_glob_warning" : Bool = PLC DB_ALARM.WRONG.rop_glob_warning AT %DB100.DBX3.6, 1 s
   "DB_ALARM_WRONG_rop_active_autocale" : Bool = PLC DB_ALARM.WRONG.rop_active_autocale AT %DB100.DBX3.7, 1 s
   "DB_ALARM_wrong_line" : Int = PLC DB_ALARM.wrong_line AT %DB100.DBW256, 1 s
   "DB_ALARM_wrong_op_1" : Int = PLC DB_ALARM.wrong_op_1 AT %DB100.DBW260, 1 s
   "DB_ALARM_wrong_op_2" : Int = PLC DB_ALARM.wrong_op_2 AT %DB100.DBW264, 1 s
   "DB_ALARM_wrong_op_3" : Int = PLC DB_ALARM.wrong_op_3 AT %DB100.DBW268, 1 s
   "DB_ALARM_alarm_line" : Int = PLC DB_ALARM.alarm_line AT %DB100.DBW254, 1 s
   "DB_ALARM_alarm_op_1" : Int = PLC DB_ALARM.alarm_op_1 AT %DB100.DBW258, 1 s
   "DB_ALARM_alarm_op_2" : Int = PLC DB_ALARM.alarm_op_2 AT %DB100.DBW262, 1 s
   "DB_ALARM_alarm_op_3" : Int = PLC DB_ALARM.alarm_op_3 AT %DB100.DBW266, 1 s
   "DB_ALARM_alarm_op_4" : Int = PLC DB_ALARM.alarm_op_4 AT %DB100.DBW270, 1 s

discrete alarms
   96: 'op_2_wrong_16', class warning_individual, trigger "DB_ALARM_wrong_op_2" bit 15
   95: 'op_2_wrong_15', class warning_individual, trigger "DB_ALARM_wrong_op_2" bit 14
   114: 'op_3_wrong_2', class warning_individual, trigger "DB_ALARM_wrong_op_3" bit 1
   113: 'op_3_wrong_1', class warning_individual, trigger "DB_ALARM_wrong_op_3" bit 0
   93: 'op_2_wrong_13', class warning_individual, trigger "DB_ALARM_wrong_op_2" bit 12
   30: 'wrong_line_14', class warning_individual, trigger "DB_ALARM_wrong_line" bit 13
   31: 'Zařízení ropex není ve standartním stavu otevřete obrazovku ROPEX + PODÉLNÉ ČELISTI a zkontorlujte hlášení', class warning_individual, trigger "DB_ALARM_wrong_line" bit 14
   32: 'Ropex provádí kalibraci vyčkejte (ROPEX + PODÉLNÉ ČELISTI)', class warning_individual, trigger "DB_ALARM_wrong_line" bit 15
   90: 'op_2_wrong_10', class warning_individual, trigger "DB_ALARM_wrong_op_2" bit 9
   89: 'op_2_wrong_9', class warning_individual, trigger "DB_ALARM_wrong_op_2" bit 8
   49: 'op_1_wrong_1', class warning_individual, trigger "DB_ALARM_wrong_op_1" bit 0
   50: 'op_1_wrong_2', class warning_individual, trigger "DB_ALARM_wrong_op_1" bit 1
   51: 'op_1_wrong_3', class warning_individual, trigger "DB_ALARM_wrong_op_1" bit 2
   52: 'op_1_wrong_4', class warning_individual, trigger "DB_ALARM_wrong_op_1" bit 3
   53: 'op_1_wrong_5', class warning_individual, trigger "DB_ALARM_wrong_op_1" bit 4
   54: 'op_1_wrong_6', class warning_individual, trigger "DB_ALARM_wrong_op_1" bit 5
   55: 'op_1_wrong_7', class warning_individual, trigger "DB_ALARM_wrong_op_1" bit 6
   56: 'op_1_wrong_8', class warning_individual, trigger "DB_ALARM_wrong_op_1" bit 7
   57: 'op_1_wrong_9', class warning_individual, trigger "DB_ALARM_wrong_op_1" bit 8
   58: 'op_1_wrong_10', class warning_individual, trigger "DB_ALARM_wrong_op_1" bit 9
   59: 'op_1_wrong_11', class warning_individual, trigger "DB_ALARM_wrong_op_1" bit 10
   60: 'op_1_wrong_12', class warning_individual, trigger "DB_ALARM_wrong_op_1" bit 11
   61: 'op_1_wrong_13', class warning_individual, trigger "DB_ALARM_wrong_op_1" bit 12
   62: 'op_1_wrong_14', class warning_individual, trigger "DB_ALARM_wrong_op_1" bit 13
   63: 'op_1_wrong_15', class warning_individual, trigger "DB_ALARM_wrong_op_1" bit 14
   64: 'op_1_wrong_16', class warning_individual, trigger "DB_ALARM_wrong_op_1" bit 15
   88: 'op_2_wrong_8', class warning_individual, trigger "DB_ALARM_wrong_op_2" bit 7
   87: 'op_2_wrong_7', class warning_individual, trigger "DB_ALARM_wrong_op_2" bit 6
   81: 'op_2_wrong_1', class warning_individual, trigger "DB_ALARM_wrong_op_2" bit 0
   82: 'op_2_wrong_2', class warning_individual, trigger "DB_ALARM_wrong_op_2" bit 1
   83: 'op_2_wrong_3', class warning_individual, trigger "DB_ALARM_wrong_op_2" bit 2
   84: 'op_2_wrong_4', class warning_individual, trigger "DB_ALARM_wrong_op_2" bit 3
   29: 'wrong_line_13', class warning_individual, trigger "DB_ALARM_wrong_line" bit 12
   94: 'op_2_wrong_14', class warning_individual, trigger "DB_ALARM_wrong_op_2" bit 13
   28: 'wrong_line_12', class warning_individual, trigger "DB_ALARM_wrong_line" bit 11
   26: 'Globální upozornění - zařízení nebo část není ve standardu', class warning_individual, trigger "DB_ALARM_wrong_line" bit 9
   92: 'op_2_wrong_12', class warning_individual, trigger "DB_ALARM_wrong_op_2" bit 11
   91: 'op_2_wrong_11', class warning_individual, trigger "DB_ALARM_wrong_op_2" bit 10
   17: 'wrong_line_1', class warning_individual, trigger "DB_ALARM_wrong_line" bit 0
   18: 'wrong_line_2', class warning_individual, trigger "DB_ALARM_wrong_line" bit 1
   19: 'wrong_line_3', class warning_individual, trigger "DB_ALARM_wrong_line" bit 2
   20: 'wrong_line_4', class warning_individual, trigger "DB_ALARM_wrong_line" bit 3
   21: 'wrong_line_5', class warning_individual, trigger "DB_ALARM_wrong_line" bit 4
   22: 'wrong_line_6', class warning_individual, trigger "DB_ALARM_wrong_line" bit 5
   23: 'Čelisti ropex je nutné zkontrolovat', class warning_individual, trigger "DB_ALARM_wrong_line" bit 6
   24: 'Ropex autocal aktivní', class warning_individual, trigger "DB_ALARM_wrong_line" bit 7
   25: 'Běží inicializace VYČKEJTE', class warning_individual, trigger "DB_ALARM_wrong_line" bit 8
   27: 'wrong_line_11', class warning_individual, trigger "DB_ALARM_wrong_line" bit 10
   45: 'op_1_alrm_13', class Errors, trigger "DB_ALARM_alarm_op_1" bit 12
   46: 'op_1_alrm_14', class Errors, trigger "DB_ALARM_alarm_op_1" bit 13
   47: 'op_1_alrm_15', class Errors, trigger "DB_ALARM_alarm_op_1" bit 14
   48: 'Měření hladiny tužek - senzro je v poruše zkontrolujte / srovnejte hladinu tužek', class Errors, trigger "DB_ALARM_alarm_op_1" bit 15
   124: 'op_3_wrong_12', class warning_individual, trigger "DB_ALARM_wrong_op_3" bit 11
   123: 'op_3_wrong_11', class warning_individual, trigger "DB_ALARM_wrong_op_3" bit 10
   65: 'SERVO SELHÁNÍ BLOKU OVLÁDÁNÍ "JOG"( KONTAKTUJTE LIFTEC)', class Errors, trigger "DB_ALARM_alarm_op_2" bit 0
   66: 'SERVO - NEZDAŘIL SE RESET N-CODÉRU - PŘEPNĚTE DO MANULÁLU A ZPĚT', class Errors, trigger "DB_ALARM_alarm_op_2" bit 1
   67: 'NEDOVŘENÍ PODÉLNÝCH ČELISTÍ -17B2 - (zkontrolujte prostor Čelistí a spusťte výrobu)', class Errors, trigger "DB_ALARM_alarm_op_2" bit 2
   68: 'PŘEKROČENÍ HLADINY -20B20 ZKONTROLUJTE ZDA NEPROJELI DVĚ TUŽKY NA SOBĚ / ZKŘÍPNUTÍ TUŽKY POD SEGMENTEM !', class Errors, trigger "DB_ALARM_alarm_op_2" bit 3
   69: 'op_2_alrm_5', class Errors, trigger "DB_ALARM_alarm_op_2" bit 4
   70: 'op_2_alrm_6', class Errors, trigger "DB_ALARM_alarm_op_2" bit 5
   71: 'DOŠLA FOLIE -21B3', class Errors, trigger "DB_ALARM_alarm_op_2" bit 6
   72: 'op_2_alrm_8', class Errors, trigger "DB_ALARM_alarm_op_2" bit 7
   73: 'OTEVŘEN BEZPEČNOSTNÍ KRYT (dveře 1)', class Errors, trigger "DB_ALARM_alarm_op_2" bit 8
   74: 'OTEVŘEN BEZPEČNOSTNÍ KRYT (dveře 2)', class Errors, trigger "DB_ALARM_alarm_op_2" bit 9
   75: 'OTEVŘEN BEZPEČNOSTNÍ KRYT (dveře 3)', class Errors, trigger "DB_ALARM_alarm_op_2" bit 10
   76: 'OTEVŘEN BEZPEČNOSTNÍ KRYT (dveře 4)', class Errors, trigger "DB_ALARM_alarm_op_2" bit 11
   77: 'PŘERUŠEN BEZPEČNOSTNÍ PAPRSEK V TUNELU', class Errors, trigger "DB_ALARM_alarm_op_2" bit 12
   78: 'PORUCHA ROPEXU PROVEĎTE INICIALIZACI ( PŘEPNUTÍM REŽIMŮ)', class Errors, trigger "DB_ALARM_alarm_op_2" bit 13
   79: 'ROPEX ALARM ZKONTROLUJTE OBRAZOVKU (ROPEX + PODÉLNÉ ČELISTI)', class Errors, trigger "DB_ALARM_alarm_op_2" bit 14
   80: 'SERVO SELHÁNÍ BLOKU OVLÁDÁNÍ "POWER" (KONTAKTUJTE LIFTEC)', class Errors, trigger "DB_ALARM_alarm_op_2" bit 15
   122: 'op_3_wrong_10', class warning_individual, trigger "DB_ALARM_wrong_op_3" bit 9
   121: 'op_3_wrong_9', class warning_individual, trigger "DB_ALARM_wrong_op_3" bit 8
   97: 'op_3_alarm_1', class Errors, trigger "DB_ALARM_alarm_op_3" bit 0
   98: 'op_3_alarm_2', class Errors, trigger "DB_ALARM_alarm_op_3" bit 1
   99: 'op_3_alarm_3', class Errors, trigger "DB_ALARM_alarm_op_3" bit 2
   44: 'op_1_alrm_12', class Errors, trigger "DB_ALARM_alarm_op_1" bit 11
   43: 'op_1_alrm_11', class Errors, trigger "DB_ALARM_alarm_op_1" bit 10
   42: 'op_1_alrm_10', class Errors, trigger "DB_ALARM_alarm_op_1" bit 9
   41: 'OTEVŘEN BEZPEČNOSTNÍ KRYT (dveře 1)', class Errors, trigger "DB_ALARM_alarm_op_1" bit 8
   128: 'op_3_wrong_16', class warning_individual, trigger "DB_ALARM_wrong_op_3" bit 15
   127: 'op_3_wrong_15', class warning_individual, trigger "DB_ALARM_wrong_op_3" bit 14
   1: 'Tiskárna nekomunikuje', class Errors, trigger "DB_ALARM_alarm_line" bit 0
   2: 'Boční kamera L offline', class Errors, trigger "DB_ALARM_alarm_line" bit 1
   3: 'Boční kamera P offline', class Errors, trigger "DB_ALARM_alarm_line" bit 2
   4: 'Horní kamera (etiketa) offline', class Errors, trigger "DB_ALARM_alarm_line" bit 3
   5: 'Chybné datum v receptuře – tiskne se XX.XX.XXXX', class Errors, trigger "DB_ALARM_alarm_line" bit 4
   6: 'Fronta plná – výsledky se nezapisují, resetujte frontu', class Errors, trigger "DB_ALARM_alarm_line" bit 5
   7: 'Horní kamera: job se nepodařilo načíst', class Errors, trigger "DB_ALARM_alarm_line" bit 6
   8: 'Otevřené levé dveře', class Errors, trigger "DB_ALARM_alarm_line" bit 7
   9: 'Otevřené pravé dveře', class Errors, trigger "DB_ALARM_alarm_line" bit 8
   10: 'APLIKÁTOR ETIKET V PORUŠE ZKONTROLUJTE', class Errors, trigger "DB_ALARM_alarm_line" bit 9
   11: 'alarm_line_11', class Errors, trigger "DB_ALARM_alarm_line" bit 10
   100: 'op_3_alarm_4', class Errors, trigger "DB_ALARM_alarm_op_3" bit 3
   12: 'alarm_line_12', class Errors, trigger "DB_ALARM_alarm_line" bit 11
   14: 'alarm_line_14', class Errors, trigger "DB_ALARM_alarm_line" bit 13
   15: 'Nedostatečný tlak vzduchu', class Errors, trigger "DB_ALARM_alarm_line" bit 14
   16: 'alarm_line_16', class Errors, trigger "DB_ALARM_alarm_line" bit 15
   126: 'op_3_wrong_14', class warning_individual, trigger "DB_ALARM_wrong_op_3" bit 13
   125: 'op_3_wrong_13', class warning_individual, trigger "DB_ALARM_wrong_op_3" bit 12
   33: 'op_1_alrm_1', class Errors, trigger "DB_ALARM_alarm_op_1" bit 0
   34: 'op_1_alrm_2', class Errors, trigger "DB_ALARM_alarm_op_1" bit 1
   35: 'op_1_alrm_3', class Errors, trigger "DB_ALARM_alarm_op_1" bit 2
   36: 'op_1_alrm_4', class Errors, trigger "DB_ALARM_alarm_op_1" bit 3
   37: 'op_1_alrm_5', class Errors, trigger "DB_ALARM_alarm_op_1" bit 4
   38: 'op_1_alrm_6', class Errors, trigger "DB_ALARM_alarm_op_1" bit 5
   39: 'op_1_alrm_7', class Errors, trigger "DB_ALARM_alarm_op_1" bit 6
   40: 'op_1_alrm_8', class Errors, trigger "DB_ALARM_alarm_op_1" bit 7
   13: 'alarm_line_13', class Errors, trigger "DB_ALARM_alarm_line" bit 12
   101: 'op_3_alarm_5', class Errors, trigger "DB_ALARM_alarm_op_3" bit 4
   103: 'op_3_alarm_7', class Errors, trigger "DB_ALARM_alarm_op_3" bit 6
   163: 'OP1_N0 -Y7 Externí alarm err 2', class Errors, trigger "DB_ALARM_OP1_M_0" bit 2
   164: 'OP1_N0 -Y7 Externí alarm err 3', class Errors, trigger "DB_ALARM_OP1_M_0" bit 3
   165: 'OP1_N0 -Y7 Motor nemá splněny podmínky pro opuštění pozice HOME', class Errors, trigger "DB_ALARM_OP1_M_0" bit 4
   166: 'OP1_N0 -Y7 Motor nemá splněny podmínky pro opuštění pozice WORK', class Errors, trigger "DB_ALARM_OP1_M_0" bit 5
   167: 'OP1_N0 -Y7 Motor nedojel do požadované pozice WORK', class Errors, trigger "DB_ALARM_OP1_M_0" bit 6
   168: 'OP1_N0 -Y7 Motor nedojel do požadované pozice HOME', class Errors, trigger "DB_ALARM_OP1_M_0" bit 7
   169: 'OP1_-Y7 RESERVE_1', class Errors, trigger "DB_ALARM_OP1_M_0" bit 8
   170: 'OP1_-Y7 RESERVE_2', class Errors, trigger "DB_ALARM_OP1_M_0" bit 9
   171: 'OP1_-Y7 RESERVE_3', class Errors, trigger "DB_ALARM_OP1_M_0" bit 10
   172: 'OP1_-Y7 RESERVE_4', class Errors, trigger "DB_ALARM_OP1_M_0" bit 11
   173: 'OP1_-Y7 RESERVE_5', class Errors, trigger "DB_ALARM_OP1_M_0" bit 12
   174: 'OP1_-Y7 RESERVE_6', class Errors, trigger "DB_ALARM_OP1_M_0" bit 13
   175: 'OP1_-Y7 RESERVE_7', class Errors, trigger "DB_ALARM_OP1_M_0" bit 14
   176: 'OP1_-Y7 RESERVE_8', class Errors, trigger "DB_ALARM_OP1_M_0" bit 15
   116: 'op_3_wrong_4', class warning_individual, trigger "DB_ALARM_wrong_op_3" bit 3
   115: 'op_3_wrong_3', class warning_individual, trigger "DB_ALARM_wrong_op_3" bit 2
   85: 'op_2_wrong_5', class warning_individual, trigger "DB_ALARM_wrong_op_2" bit 4
   162: 'OP1_N0 -Y7 Externí alarm err 1', class Errors, trigger "DB_ALARM_OP1_M_0" bit 1
   102: 'op_3_alarm_6', class Errors, trigger "DB_ALARM_alarm_op_3" bit 5
   161: 'OP1_N0 -Y7 Nespecifikovaný režim motoru AUTOMAT/MANUAL', class Errors, trigger "DB_ALARM_OP1_M_0" bit 0
   118: 'op_3_wrong_6', class warning_individual, trigger "DB_ALARM_wrong_op_3" bit 5
   104: 'op_3_alarm_8', class Errors, trigger "DB_ALARM_alarm_op_3" bit 7
   105: 'op_3_alarm_9', class Errors, trigger "DB_ALARM_alarm_op_3" bit 8
   106: 'op_3_alarm_10', class Errors, trigger "DB_ALARM_alarm_op_3" bit 9
   107: 'op_3_alarm_11', class Errors, trigger "DB_ALARM_alarm_op_3" bit 10
   108: 'op_3_alarm_12', class Errors, trigger "DB_ALARM_alarm_op_3" bit 11
   109: 'op_3_alarm_13', class Errors, trigger "DB_ALARM_alarm_op_3" bit 12
   110: 'op_3_alarm_14', class Errors, trigger "DB_ALARM_alarm_op_3" bit 13
   111: 'op_3_alarm_15', class Errors, trigger "DB_ALARM_alarm_op_3" bit 14
   112: 'op_3_alarm_16', class Errors, trigger "DB_ALARM_alarm_op_3" bit 15
   120: 'op_3_wrong_8', class warning_individual, trigger "DB_ALARM_wrong_op_3" bit 7
   119: 'op_3_wrong_7', class warning_individual, trigger "DB_ALARM_wrong_op_3" bit 6
   145: 'OP0_N0 Nespecifikovaný režim motoru AUTOMAT/MANUAL', class Errors bit 0
   146: 'OP0_N0 Externí alarm err 1', class Errors bit 0
   117: 'op_3_wrong_5', class warning_individual, trigger "DB_ALARM_wrong_op_3" bit 4
   147: 'OP0_N0 Externí alarm err 2', class Errors bit 0
   149: 'OP0_N0 Motor nemá splněny podmínky pro opuštění pozice HOME', class Errors bit 0
   150: 'OP0_N0 Motor nemá splněny podmínky pro opuštění pozice WORK', class Errors bit 0
   151: 'OP0_N0 Motor nedojel do požadované pozice WORK', class Errors bit 0
   152: 'OP0_N0 Motor nedojel do požadované pozice HOME', class Errors bit 0
   153: 'op_0_m_0_8', class Errors bit 0
   154: 'op_0_m_0_9', class Errors bit 0
   155: 'op_0_m_0_10', class Errors bit 0
   156: 'op_0_m_0_11', class Errors bit 0
   157: 'op_0_m_0_12', class Errors bit 0
   158: 'op_0_m_0_13', class Errors bit 0
   159: 'op_0_m_0_14', class Errors bit 0
   160: 'op_0_m_0_15', class Errors bit 0
   148: 'OP0_N0 Externí alarm err 3', class Errors bit 0
   86: 'op_2_wrong_6', class warning_individual, trigger "DB_ALARM_wrong_op_2" bit 5
   177: 'OP1_N0 -Y9 Nespecifikovaný režim motoru AUTOMAT/MANUAL', class Errors, trigger "DB_ALARM_OP1_M_1" bit 0
   178: 'OP1_N0 -Y9 Externí alarm err 1', class Errors, trigger "DB_ALARM_OP1_M_1" bit 1
   179: 'OP1_N0 -Y9 Externí alarm err 2', class Errors, trigger "DB_ALARM_OP1_M_1" bit 2
   180: 'OP1_N0 -Y9 Externí alarm err 3', class Errors, trigger "DB_ALARM_OP1_M_1" bit 3
   181: 'OP1_N0 -Y9 Motor nemá splněny podmínky pro opuštění pozice HOME', class Errors, trigger "DB_ALARM_OP1_M_1" bit 4
   182: 'OP1_N0 -Y9 Motor nemá splněny podmínky pro opuštění pozice WORK', class Errors, trigger "DB_ALARM_OP1_M_1" bit 5
   183: 'OP1_N0 -Y9 Motor nedojel do požadované pozice WORK', class Errors, trigger "DB_ALARM_OP1_M_1" bit 6
   184: 'OP1_N0 -Y9 Motor nedojel do požadované pozice HOME', class Errors, trigger "DB_ALARM_OP1_M_1" bit 7
   185: 'OP1_RESERVE_1 -Y9', class Errors, trigger "DB_ALARM_OP1_M_1" bit 8
   186: 'OP1_RESERVE_2 -Y9', class Errors, trigger "DB_ALARM_OP1_M_1" bit 9
   187: 'OP1_RESERVE_3 -Y9', class Errors, trigger "DB_ALARM_OP1_M_1" bit 10
   188: 'OP1_RESERVE_4 -Y9', class Errors, trigger "DB_ALARM_OP1_M_1" bit 11
   189: 'OP1_RESERVE_5 -Y9', class Errors, trigger "DB_ALARM_OP1_M_1" bit 12
   190: 'OP1_RESERVE_6 -Y9', class Errors, trigger "DB_ALARM_OP1_M_1" bit 13
   191: 'OP1_RESERVE_7 -Y9', class Errors, trigger "DB_ALARM_OP1_M_1" bit 14
   192: 'OP1_RESERVE_8 -Y9', class Errors, trigger "DB_ALARM_OP1_M_1" bit 15
   193: 'OP1_N0 Nespecifikovaný režim motoru AUTOMAT/MANUAL', class Errors, trigger "DB_ALARM_OP1_M_2" bit 0
   194: 'OP1_N0 Externí alarm err 1', class Errors, trigger "DB_ALARM_OP1_M_2" bit 1
   195: 'OP1_N0 Externí alarm err 2', class Errors, trigger "DB_ALARM_OP1_M_2" bit 2
   196: 'OP1_N0 Externí alarm err 3', class Errors, trigger "DB_ALARM_OP1_M_2" bit 3
   197: 'OP1_N0 Motor nemá splněny podmínky pro opuštění pozice HOME', class Errors, trigger "DB_ALARM_OP1_M_2" bit 4
   198: 'OP1_N0 Motor nemá splněny podmínky pro opuštění pozice WORK', class Errors, trigger "DB_ALARM_OP1_M_2" bit 5
   199: 'OP1_N0 Motor nedojel do požadované pozice WORK', class Errors, trigger "DB_ALARM_OP1_M_2" bit 6
   200: 'OP1_N0 Motor nedojel do požadované pozice HOME', class Errors, trigger "DB_ALARM_OP1_M_2" bit 7
   201: 'OP1_RESERVE_1', class Errors, trigger "DB_ALARM_OP1_M_2" bit 8
   202: 'OP1_RESERVE_2', class Errors, trigger "DB_ALARM_OP1_M_2" bit 9
   203: 'OP1_RESERVE_3', class Errors, trigger "DB_ALARM_OP1_M_2" bit 10
   204: 'OP1_RESERVE_4', class Errors, trigger "DB_ALARM_OP1_M_2" bit 11
   205: 'OP1_RESERVE_5', class Errors, trigger "DB_ALARM_OP1_M_2" bit 12
   206: 'OP1_RESERVE_6', class Errors, trigger "DB_ALARM_OP1_M_2" bit 13
   207: 'OP1_RESERVE_7', class Errors, trigger "DB_ALARM_OP1_M_2" bit 14
   208: 'OP1_RESERVE_8', class Errors, trigger "DB_ALARM_OP1_M_2" bit 15
   209: 'OP1_N0 Nespecifikovaný režim motoru AUTOMAT/MANUAL', class Errors, trigger "DB_ALARM_OP1_M_3" bit 0
   210: 'OP1_N0 Externí alarm err 1', class Errors, trigger "DB_ALARM_OP1_M_3" bit 1
   211: 'OP1_N0 Externí alarm err 2', class Errors, trigger "DB_ALARM_OP1_M_3" bit 2
   212: 'OP1_N0 Externí alarm err 3', class Errors, trigger "DB_ALARM_OP1_M_3" bit 3
   213: 'OP1_N0 Motor nemá splněny podmínky pro opuštění pozice HOME', class Errors, trigger "DB_ALARM_OP1_M_3" bit 4
   214: 'OP1_N0 Motor nemá splněny podmínky pro opuštění pozice WORK', class Errors, trigger "DB_ALARM_OP1_M_3" bit 5
   215: 'OP1_N0 Motor nedojel do požadované pozice WORK', class Errors, trigger "DB_ALARM_OP1_M_3" bit 6
   216: 'OP1_N0 Motor nedojel do požadované pozice HOME', class Errors, trigger "DB_ALARM_OP1_M_3" bit 7
   217: 'OP1_RESERVE_1', class Errors, trigger "DB_ALARM_OP1_M_3" bit 8
   218: 'OP1_RESERVE_2', class Errors, trigger "DB_ALARM_OP1_M_3" bit 9
   219: 'OP1_RESERVE_3', class Errors, trigger "DB_ALARM_OP1_M_3" bit 10
   220: 'OP1_RESERVE_4', class Errors, trigger "DB_ALARM_OP1_M_3" bit 11
   221: 'OP1_RESERVE_5', class Errors, trigger "DB_ALARM_OP1_M_3" bit 12
   222: 'OP1_RESERVE_6', class Errors, trigger "DB_ALARM_OP1_M_3" bit 13
   223: 'OP1_RESERVE_7', class Errors, trigger "DB_ALARM_OP1_M_3" bit 14
   224: 'OP1_RESERVE_8', class Errors, trigger "DB_ALARM_OP1_M_3" bit 15
   225: 'OP1_N0 Nespecifikovaný režim motoru AUTOMAT/MANUAL', class Errors, trigger "DB_ALARM_OP1_M_4" bit 0
   226: 'OP1_N0 Externí alarm err 1', class Errors, trigger "DB_ALARM_OP1_M_4" bit 1
   227: 'OP1_N0 Externí alarm err 2', class Errors, trigger "DB_ALARM_OP1_M_4" bit 2
   228: 'OP1_N0 Externí alarm err 3', class Errors, trigger "DB_ALARM_OP1_M_4" bit 3
   229: 'OP1_N0 Motor nemá splněny podmínky pro opuštění pozice HOME', class Errors, trigger "DB_ALARM_OP1_M_4" bit 4
   230: 'OP1_N0 Motor nemá splněny podmínky pro opuštění pozice WORK', class Errors, trigger "DB_ALARM_OP1_M_4" bit 5
   231: 'OP1_N0 Motor nedojel do požadované pozice WORK', class Errors, trigger "DB_ALARM_OP1_M_4" bit 6
   232: 'OP1_N0 Motor nedojel do požadované pozice HOME', class Errors, trigger "DB_ALARM_OP1_M_4" bit 7
   233: 'OP1_RESERVE_1', class Errors, trigger "DB_ALARM_OP1_M_4" bit 8
   234: 'OP1_RESERVE_2', class Errors, trigger "DB_ALARM_OP1_M_4" bit 9
   235: 'OP1_RESERVE_3', class Errors, trigger "DB_ALARM_OP1_M_4" bit 10
   236: 'OP1_RESERVE_4', class Errors, trigger "DB_ALARM_OP1_M_4" bit 11
   237: 'OP1_RESERVE_5', class Errors, trigger "DB_ALARM_OP1_M_4" bit 12
   238: 'OP1_RESERVE_6', class Errors, trigger "DB_ALARM_OP1_M_4" bit 13
   239: 'OP1_RESERVE_7', class Errors, trigger "DB_ALARM_OP1_M_4" bit 14
   240: 'OP1_RESERVE_8', class Errors, trigger "DB_ALARM_OP1_M_4" bit 15
   241: 'OP1_N0 Nespecifikovaný režim motoru AUTOMAT/MANUAL', class Errors, trigger "DB_ALARM_OP1_M_5" bit 0
   242: 'OP1_N0 Externí alarm err 1', class Errors, trigger "DB_ALARM_OP1_M_5" bit 1
   243: 'OP1_N0 Externí alarm err 2', class Errors, trigger "DB_ALARM_OP1_M_5" bit 2
   244: 'OP1_N0 Externí alarm err 3', class Errors, trigger "DB_ALARM_OP1_M_5" bit 3
   245: 'OP1_N0 Motor nemá splněny podmínky pro opuštění pozice HOME', class Errors, trigger "DB_ALARM_OP1_M_5" bit 4
   246: 'OP1_N0 Motor nemá splněny podmínky pro opuštění pozice WORK', class Errors, trigger "DB_ALARM_OP1_M_5" bit 5
   247: 'OP1_N0 Motor nedojel do požadované pozice WORK', class Errors, trigger "DB_ALARM_OP1_M_5" bit 6
   248: 'OP1_N0 Motor nedojel do požadované pozice HOME', class Errors, trigger "DB_ALARM_OP1_M_5" bit 7
   249: 'OP1_RESERVE_1', class Errors, trigger "DB_ALARM_OP1_M_5" bit 8
   250: 'OP1_RESERVE_2', class Errors, trigger "DB_ALARM_OP1_M_5" bit 9
   251: 'OP1_RESERVE_3', class Errors, trigger "DB_ALARM_OP1_M_5" bit 10
   252: 'OP1_RESERVE_4', class Errors, trigger "DB_ALARM_OP1_M_5" bit 11
   253: 'OP1_RESERVE_5', class Errors, trigger "DB_ALARM_OP1_M_5" bit 12
   254: 'OP1_RESERVE_6', class Errors, trigger "DB_ALARM_OP1_M_5" bit 13
   255: 'OP1_RESERVE_7', class Errors, trigger "DB_ALARM_OP1_M_5" bit 14
   256: 'OP1_RESERVE_8', class Errors, trigger "DB_ALARM_OP1_M_5" bit 15
   257: 'OP1_N0 Nespecifikovaný režim motoru AUTOMAT/MANUAL', class Errors, trigger "DB_ALARM_OP1_M_6" bit 0
   258: 'OP1_N0 Externí alarm err 1', class Errors, trigger "DB_ALARM_OP1_M_6" bit 1
   259: 'OP1_N0 Externí alarm err 2', class Errors, trigger "DB_ALARM_OP1_M_6" bit 2
   260: 'OP1_N0 Externí alarm err 3', class Errors, trigger "DB_ALARM_OP1_M_6" bit 3
   261: 'OP1_N0 Motor nemá splněny podmínky pro opuštění pozice HOME', class Errors, trigger "DB_ALARM_OP1_M_6" bit 4
   262: 'OP1_N0 Motor nemá splněny podmínky pro opuštění pozice WORK', class Errors, trigger "DB_ALARM_OP1_M_6" bit 5
   263: 'OP1_N0 Motor nedojel do požadované pozice WORK', class Errors, trigger "DB_ALARM_OP1_M_6" bit 6
   264: 'OP1_N0 Motor nedojel do požadované pozice HOME', class Errors, trigger "DB_ALARM_OP1_M_6" bit 7
   265: 'OP1_RESERVE_1', class Errors, trigger "DB_ALARM_OP1_M_6" bit 8
   266: 'OP1_RESERVE_2', class Errors, trigger "DB_ALARM_OP1_M_6" bit 9
   267: 'OP1_RESERVE_3', class Errors, trigger "DB_ALARM_OP1_M_6" bit 10
   268: 'OP1_RESERVE_4', class Errors, trigger "DB_ALARM_OP1_M_6" bit 11
   269: 'OP1_RESERVE_5', class Errors, trigger "DB_ALARM_OP1_M_6" bit 12
   270: 'OP1_RESERVE_6', class Errors, trigger "DB_ALARM_OP1_M_6" bit 13
   271: 'OP1_RESERVE_7', class Errors, trigger "DB_ALARM_OP1_M_6" bit 14
   272: 'OP1_RESERVE_8', class Errors, trigger "DB_ALARM_OP1_M_6" bit 15
   273: 'OP1_N0 Nespecifikovaný režim motoru AUTOMAT/MANUAL', class Errors, trigger "DB_ALARM_OP1_M_7" bit 0
   274: 'OP1_N0 Externí alarm err 1', class Errors, trigger "DB_ALARM_OP1_M_7" bit 1
   275: 'OP1_N0 Externí alarm err 2', class Errors, trigger "DB_ALARM_OP1_M_7" bit 2
   276: 'OP1_N0 Externí alarm err 3', class Errors, trigger "DB_ALARM_OP1_M_7" bit 3
   277: 'OP1_N0 Motor nemá splněny podmínky pro opuštění pozice HOME', class Errors, trigger "DB_ALARM_OP1_M_7" bit 4
   278: 'OP1_N0 Motor nemá splněny podmínky pro opuštění pozice WORK', class Errors, trigger "DB_ALARM_OP1_M_7" bit 5
   279: 'OP1_N0 Motor nedojel do požadované pozice WORK', class Errors, trigger "DB_ALARM_OP1_M_7" bit 6
   280: 'OP1_N0 Motor nedojel do požadované pozice HOME', class Errors, trigger "DB_ALARM_OP1_M_7" bit 7
   281: 'OP1_RESERVE_1', class Errors, trigger "DB_ALARM_OP1_M_7" bit 8
   282: 'OP1_RESERVE_2', class Errors, trigger "DB_ALARM_OP1_M_7" bit 9
   283: 'OP1_RESERVE_3', class Errors, trigger "DB_ALARM_OP1_M_7" bit 10
   284: 'OP1_RESERVE_4', class Errors, trigger "DB_ALARM_OP1_M_7" bit 11
   285: 'OP1_RESERVE_5', class Errors, trigger "DB_ALARM_OP1_M_7" bit 12
   286: 'OP1_RESERVE_6', class Errors, trigger "DB_ALARM_OP1_M_7" bit 13
   287: 'OP1_RESERVE_7', class Errors, trigger "DB_ALARM_OP1_M_7" bit 14
   288: 'OP1_RESERVE_8', class Errors, trigger "DB_ALARM_OP1_M_7" bit 15
   289: 'OP1_N0 Nespecifikovaný režim motoru AUTOMAT/MANUAL', class Errors, trigger "DB_ALARM_OP1_M_8" bit 0
   290: 'OP1_N0 Externí alarm err 1', class Errors, trigger "DB_ALARM_OP1_M_8" bit 1
   291: 'OP1_N0 Externí alarm err 2', class Errors, trigger "DB_ALARM_OP1_M_8" bit 2
   292: 'OP1_N0 Externí alarm err 3', class Errors, trigger "DB_ALARM_OP1_M_8" bit 3
   293: 'OP1_N0 Motor nemá splněny podmínky pro opuštění pozice HOME', class Errors, trigger "DB_ALARM_OP1_M_8" bit 4
   294: 'OP1_N0 Motor nemá splněny podmínky pro opuštění pozice WORK', class Errors, trigger "DB_ALARM_OP1_M_8" bit 5
   295: 'OP1_N0 Motor nedojel do požadované pozice WORK', class Errors, trigger "DB_ALARM_OP1_M_8" bit 6
   296: 'OP1_N0 Motor nedojel do požadované pozice HOME', class Errors, trigger "DB_ALARM_OP1_M_8" bit 7
   297: 'OP1_RESERVE_1', class Errors, trigger "DB_ALARM_OP1_M_8" bit 8
   298: 'OP1_RESERVE_2', class Errors, trigger "DB_ALARM_OP1_M_8" bit 9
   299: 'OP1_RESERVE_3', class Errors, trigger "DB_ALARM_OP1_M_8" bit 10
   300: 'OP1_RESERVE_4', class Errors, trigger "DB_ALARM_OP1_M_8" bit 11
   301: 'OP1_RESERVE_5', class Errors, trigger "DB_ALARM_OP1_M_8" bit 12
   302: 'OP1_RESERVE_6', class Errors, trigger "DB_ALARM_OP1_M_8" bit 13
   303: 'OP1_RESERVE_7', class Errors, trigger "DB_ALARM_OP1_M_8" bit 14
   304: 'OP1_RESERVE_8', class Errors, trigger "DB_ALARM_OP1_M_8" bit 15
   305: 'OP1_N0 Nespecifikovaný režim motoru AUTOMAT/MANUAL', class Errors, trigger "DB_ALARM_OP1_M_9" bit 0
   306: 'OP1_N0 Externí alarm err 1', class Errors, trigger "DB_ALARM_OP1_M_9" bit 1
   307: 'OP1_N0 Externí alarm err 2', class Errors, trigger "DB_ALARM_OP1_M_9" bit 2
   308: 'OP1_N0 Externí alarm err 3', class Errors, trigger "DB_ALARM_OP1_M_9" bit 3
   309: 'OP1_N0 Motor nemá splněny podmínky pro opuštění pozice HOME', class Errors, trigger "DB_ALARM_OP1_M_9" bit 4
   310: 'OP1_N0 Motor nemá splněny podmínky pro opuštění pozice WORK', class Errors, trigger "DB_ALARM_OP1_M_9" bit 5
   311: 'OP1_N0 Motor nedojel do požadované pozice WORK', class Errors, trigger "DB_ALARM_OP1_M_9" bit 6
   312: 'OP1_N0 Motor nedojel do požadované pozice HOME', class Errors, trigger "DB_ALARM_OP1_M_9" bit 7
   313: 'OP1_RESERVE_1', class Errors, trigger "DB_ALARM_OP1_M_9" bit 8
   314: 'OP1_RESERVE_2', class Errors, trigger "DB_ALARM_OP1_M_9" bit 9
   315: 'OP1_RESERVE_3', class Errors, trigger "DB_ALARM_OP1_M_9" bit 10
   316: 'OP1_RESERVE_4', class Errors, trigger "DB_ALARM_OP1_M_9" bit 11
   317: 'OP1_RESERVE_5', class Errors, trigger "DB_ALARM_OP1_M_9" bit 12
   318: 'OP1_RESERVE_6', class Errors, trigger "DB_ALARM_OP1_M_9" bit 13
   319: 'OP1_RESERVE_7', class Errors, trigger "DB_ALARM_OP1_M_9" bit 14
   320: 'OP1_RESERVE_8', class Errors, trigger "DB_ALARM_OP1_M_9" bit 15
   321: 'OP1_N0 Nespecifikovaný režim motoru AUTOMAT/MANUAL', class Errors, trigger "DB_ALARM_OP1_M_10" bit 0
   322: 'OP1_N0 Externí alarm err 1', class Errors, trigger "DB_ALARM_OP1_M_10" bit 1
   323: 'OP1_N0 Externí alarm err 2', class Errors, trigger "DB_ALARM_OP1_M_10" bit 2
   324: 'OP1_N0 Externí alarm err 3', class Errors, trigger "DB_ALARM_OP1_M_10" bit 3
   325: 'OP1_N0 Motor nemá splněny podmínky pro opuštění pozice HOME', class Errors, trigger "DB_ALARM_OP1_M_10" bit 4
   326: 'OP1_N0 Motor nemá splněny podmínky pro opuštění pozice WORK', class Errors, trigger "DB_ALARM_OP1_M_10" bit 5
   327: 'OP1_N0 Motor nedojel do požadované pozice WORK', class Errors, trigger "DB_ALARM_OP1_M_10" bit 6
   328: 'OP1_N0 Motor nedojel do požadované pozice HOME', class Errors, trigger "DB_ALARM_OP1_M_10" bit 7
   329: 'OP1_RESERVE_1', class Errors, trigger "DB_ALARM_OP1_M_10" bit 8
   330: 'OP1_RESERVE_2', class Errors, trigger "DB_ALARM_OP1_M_10" bit 9
   331: 'OP1_RESERVE_3', class Errors, trigger "DB_ALARM_OP1_M_10" bit 10
   332: 'OP1_RESERVE_4', class Errors, trigger "DB_ALARM_OP1_M_10" bit 11
   333: 'OP1_RESERVE_5', class Errors, trigger "DB_ALARM_OP1_M_10" bit 12
   334: 'OP1_RESERVE_6', class Errors, trigger "DB_ALARM_OP1_M_10" bit 13
   335: 'OP1_RESERVE_7', class Errors, trigger "DB_ALARM_OP1_M_10" bit 14
   336: 'OP1_RESERVE_8', class Errors, trigger "DB_ALARM_OP1_M_10" bit 15
   337: 'OP1_N0 Nespecifikovaný režim motoru AUTOMAT/MANUAL', class Errors, trigger "DB_ALARM_OP1_M_11" bit 0
   338: 'OP1_N0 Externí alarm err 1', class Errors, trigger "DB_ALARM_OP1_M_11" bit 1
   339: 'OP1_N0 Externí alarm err 2', class Errors, trigger "DB_ALARM_OP1_M_11" bit 2
   340: 'OP1_N0 Externí alarm err 3', class Errors, trigger "DB_ALARM_OP1_M_11" bit 3
   341: 'OP1_N0 Motor nemá splněny podmínky pro opuštění pozice HOME', class Errors, trigger "DB_ALARM_OP1_M_11" bit 4
   342: 'OP1_N0 Motor nemá splněny podmínky pro opuštění pozice WORK', class Errors, trigger "DB_ALARM_OP1_M_11" bit 5
   343: 'OP1_N0 Motor nedojel do požadované pozice WORK', class Errors, trigger "DB_ALARM_OP1_M_11" bit 6
   344: 'OP1_N0 Motor nedojel do požadované pozice HOME', class Errors, trigger "DB_ALARM_OP1_M_11" bit 7
   345: 'OP1_RESERVE_1', class Errors, trigger "DB_ALARM_OP1_M_11" bit 8
   346: 'OP1_RESERVE_2', class Errors, trigger "DB_ALARM_OP1_M_11" bit 9
   347: 'OP1_RESERVE_3', class Errors, trigger "DB_ALARM_OP1_M_11" bit 10
   348: 'OP1_RESERVE_4', class Errors, trigger "DB_ALARM_OP1_M_11" bit 11
   349: 'OP1_RESERVE_5', class Errors, trigger "DB_ALARM_OP1_M_11" bit 12
   350: 'OP1_RESERVE_6', class Errors, trigger "DB_ALARM_OP1_M_11" bit 13
   351: 'OP1_RESERVE_7', class Errors, trigger "DB_ALARM_OP1_M_11" bit 14
   352: 'OP1_RESERVE_8', class Errors, trigger "DB_ALARM_OP1_M_11" bit 15
   353: 'OP1_N0 Nespecifikovaný režim motoru AUTOMAT/MANUAL', class Errors, trigger "DB_ALARM_OP1_M_12" bit 0
   354: 'OP1_N0 Externí alarm err 1', class Errors, trigger "DB_ALARM_OP1_M_12" bit 1
   355: 'OP1_N0 Externí alarm err 2', class Errors, trigger "DB_ALARM_OP1_M_12" bit 2
   356: 'OP1_N0 Externí alarm err 3', class Errors, trigger "DB_ALARM_OP1_M_12" bit 3
   357: 'OP1_N0 Motor nemá splněny podmínky pro opuštění pozice HOME', class Errors, trigger "DB_ALARM_OP1_M_12" bit 4
   358: 'OP1_N0 Motor nemá splněny podmínky pro opuštění pozice WORK', class Errors, trigger "DB_ALARM_OP1_M_12" bit 5
   359: 'OP1_N0 Motor nedojel do požadované pozice WORK', class Errors, trigger "DB_ALARM_OP1_M_12" bit 6
   360: 'OP1_N0 Motor nedojel do požadované pozice HOME', class Errors, trigger "DB_ALARM_OP1_M_12" bit 7
   361: 'OP1_RESERVE_1', class Errors, trigger "DB_ALARM_OP1_M_12" bit 8
   362: 'OP1_RESERVE_2', class Errors, trigger "DB_ALARM_OP1_M_12" bit 9
   363: 'OP1_RESERVE_3', class Errors, trigger "DB_ALARM_OP1_M_12" bit 10
   364: 'OP1_RESERVE_4', class Errors, trigger "DB_ALARM_OP1_M_12" bit 11
   365: 'OP1_RESERVE_5', class Errors, trigger "DB_ALARM_OP1_M_12" bit 12
   366: 'OP1_RESERVE_6', class Errors, trigger "DB_ALARM_OP1_M_12" bit 13
   367: 'OP1_RESERVE_7', class Errors, trigger "DB_ALARM_OP1_M_12" bit 14
   368: 'OP1_RESERVE_8', class Errors, trigger "DB_ALARM_OP1_M_12" bit 15
   369: 'OP1_N0 Nespecifikovaný režim motoru AUTOMAT/MANUAL', class Errors, trigger "DB_ALARM_OP1_M_13" bit 0
   370: 'OP1_N0 Externí alarm err 1', class Errors, trigger "DB_ALARM_OP1_M_13" bit 1
   371: 'OP1_N0 Externí alarm err 2', class Errors, trigger "DB_ALARM_OP1_M_13" bit 2
   372: 'OP1_N0 Externí alarm err 3', class Errors, trigger "DB_ALARM_OP1_M_13" bit 3
   373: 'OP1_N0 Motor nemá splněny podmínky pro opuštění pozice HOME', class Errors, trigger "DB_ALARM_OP1_M_13" bit 4
   374: 'OP1_N0 Motor nemá splněny podmínky pro opuštění pozice WORK', class Errors, trigger "DB_ALARM_OP1_M_13" bit 5
   375: 'OP1_N0 Motor nedojel do požadované pozice WORK', class Errors, trigger "DB_ALARM_OP1_M_13" bit 6
   376: 'OP1_N0 Motor nedojel do požadované pozice HOME', class Errors, trigger "DB_ALARM_OP1_M_13" bit 7
   377: 'OP1_RESERVE_1', class Errors, trigger "DB_ALARM_OP1_M_13" bit 8
   378: 'OP1_RESERVE_2', class Errors, trigger "DB_ALARM_OP1_M_13" bit 9
   379: 'OP1_RESERVE_3', class Errors, trigger "DB_ALARM_OP1_M_13" bit 10
   380: 'OP1_RESERVE_4', class Errors, trigger "DB_ALARM_OP1_M_13" bit 11
   381: 'OP1_RESERVE_5', class Errors, trigger "DB_ALARM_OP1_M_13" bit 12
   382: 'OP1_RESERVE_6', class Errors, trigger "DB_ALARM_OP1_M_13" bit 13
   383: 'OP1_RESERVE_7', class Errors, trigger "DB_ALARM_OP1_M_13" bit 14
   384: 'OP1_RESERVE_8', class Errors, trigger "DB_ALARM_OP1_M_13" bit 15
   385: 'OP1_N0 Nespecifikovaný režim motoru AUTOMAT/MANUAL', class Errors, trigger "DB_ALARM_OP1_M_14" bit 0
   386: 'OP1_N0 Externí alarm err 1', class Errors, trigger "DB_ALARM_OP1_M_14" bit 1
   387: 'OP1_N0 Externí alarm err 2', class Errors, trigger "DB_ALARM_OP1_M_14" bit 2
   388: 'OP1_N0 Externí alarm err 3', class Errors, trigger "DB_ALARM_OP1_M_14" bit 3
   389: 'OP1_N0 Motor nemá splněny podmínky pro opuštění pozice HOME', class Errors, trigger "DB_ALARM_OP1_M_14" bit 4
   390: 'OP1_N0 Motor nemá splněny podmínky pro opuštění pozice WORK', class Errors, trigger "DB_ALARM_OP1_M_14" bit 5
   391: 'OP1_N0 Motor nedojel do požadované pozice WORK', class Errors, trigger "DB_ALARM_OP1_M_14" bit 6
   392: 'OP1_N0 Motor nedojel do požadované pozice HOME', class Errors, trigger "DB_ALARM_OP1_M_14" bit 7
   393: 'OP1_RESERVE_1', class Errors, trigger "DB_ALARM_OP1_M_14" bit 8
   394: 'OP1_RESERVE_2', class Errors, trigger "DB_ALARM_OP1_M_14" bit 9
   395: 'OP1_RESERVE_3', class Errors, trigger "DB_ALARM_OP1_M_14" bit 10
   396: 'OP1_RESERVE_4', class Errors, trigger "DB_ALARM_OP1_M_14" bit 11
   397: 'OP1_RESERVE_5', class Errors, trigger "DB_ALARM_OP1_M_14" bit 12
   398: 'OP1_RESERVE_6', class Errors, trigger "DB_ALARM_OP1_M_14" bit 13
   399: 'OP1_RESERVE_7', class Errors, trigger "DB_ALARM_OP1_M_14" bit 14
   400: 'OP1_RESERVE_8', class Errors, trigger "DB_ALARM_OP1_M_14" bit 15
   401: 'OP1_N0 Nespecifikovaný režim motoru AUTOMAT/MANUAL', class Errors, trigger "DB_ALARM_OP1_M_15" bit 0
   402: 'OP1_N0 Externí alarm err 1', class Errors, trigger "DB_ALARM_OP1_M_15" bit 1
   403: 'OP1_N0 Externí alarm err 2', class Errors, trigger "DB_ALARM_OP1_M_15" bit 2
   404: 'OP1_N0 Externí alarm err 3', class Errors, trigger "DB_ALARM_OP1_M_15" bit 3
   405: 'OP1_N0 Motor nemá splněny podmínky pro opuštění pozice HOME', class Errors, trigger "DB_ALARM_OP1_M_15" bit 4
   406: 'OP1_N0 Motor nemá splněny podmínky pro opuštění pozice WORK', class Errors, trigger "DB_ALARM_OP1_M_15" bit 5
   407: 'OP1_N0 Motor nedojel do požadované pozice WORK', class Errors, trigger "DB_ALARM_OP1_M_15" bit 6
   408: 'OP1_N0 Motor nedojel do požadované pozice HOME', class Errors, trigger "DB_ALARM_OP1_M_15" bit 7
   409: 'OP1_RESERVE_1', class Errors, trigger "DB_ALARM_OP1_M_15" bit 8
   410: 'OP1_RESERVE_2', class Errors, trigger "DB_ALARM_OP1_M_15" bit 9
   411: 'OP1_RESERVE_3', class Errors, trigger "DB_ALARM_OP1_M_15" bit 10
   412: 'OP1_RESERVE_4', class Errors, trigger "DB_ALARM_OP1_M_15" bit 11
   413: 'OP1_RESERVE_5', class Errors, trigger "DB_ALARM_OP1_M_15" bit 12
   414: 'OP1_RESERVE_6', class Errors, trigger "DB_ALARM_OP1_M_15" bit 13
   415: 'OP1_RESERVE_7', class Errors, trigger "DB_ALARM_OP1_M_15" bit 14
   416: 'OP1_RESERVE_8', class Errors, trigger "DB_ALARM_OP1_M_15" bit 15
   417: 'OP2_N0 -YA1 Nespecifikovaný režim motoru AUTOMAT/MANUAL', class Errors, trigger "DB_ALARM_OP2_M_0" bit 0
   418: 'OP2_N0 -YA1 Externí alarm err 1', class Errors, trigger "DB_ALARM_OP2_M_0" bit 1
   419: 'OP2_N0 -YA1 Externí alarm err 2', class Errors, trigger "DB_ALARM_OP2_M_0" bit 2
   420: 'OP2_N0 -YA1 Externí alarm err 3', class Errors, trigger "DB_ALARM_OP2_M_0" bit 3
   421: 'OP2_N0 -YA1 Motor nemá splněny podmínky pro opuštění pozice HOME', class Errors, trigger "DB_ALARM_OP2_M_0" bit 4
   422: 'OP2_N0 -YA1 Motor nemá splněny podmínky pro opuštění pozice WORK', class Errors, trigger "DB_ALARM_OP2_M_0" bit 5
   423: 'OP2_N0 -YA1 Motor nedojel do požadované pozice WORK', class Errors, trigger "DB_ALARM_OP2_M_0" bit 6
   424: 'OP2_N0 -YA1 Motor nedojel do požadované pozice HOME', class Errors, trigger "DB_ALARM_OP2_M_0" bit 7
   425: 'OP2_RESERVE_1 -YA1', class Errors, trigger "DB_ALARM_OP2_M_0" bit 8
   426: 'OP2_RESERVE_2 -YA1', class Errors, trigger "DB_ALARM_OP2_M_0" bit 9
   427: 'OP2_RESERVE_3 -YA1', class Errors, trigger "DB_ALARM_OP2_M_0" bit 10
   428: 'OP2_RESERVE_4 -YA1', class Errors, trigger "DB_ALARM_OP2_M_0" bit 11
   429: 'OP2_RESERVE_5 -YA1', class Errors, trigger "DB_ALARM_OP2_M_0" bit 12
   430: 'OP2_RESERVE_6 -YA1', class Errors, trigger "DB_ALARM_OP2_M_0" bit 13
   431: 'OP2_RESERVE_7 -YA1', class Errors, trigger "DB_ALARM_OP2_M_0" bit 14
   432: 'OP2_RESERVE_8 -YA1', class Errors, trigger "DB_ALARM_OP2_M_0" bit 15
   433: 'OP2_N0 -YA2 Nespecifikovaný režim motoru AUTOMAT/MANUAL', class Errors, trigger "DB_ALARM_OP2_M_1" bit 0
   434: 'OP2_N0 -YA2 Externí alarm err 1', class Errors, trigger "DB_ALARM_OP2_M_1" bit 1
   435: 'OP2_N0 -YA2 Externí alarm err 2', class Errors, trigger "DB_ALARM_OP2_M_1" bit 2
   436: 'OP2_N0 -YA2 Externí alarm err 3', class Errors, trigger "DB_ALARM_OP2_M_1" bit 3
   437: 'OP2_N0 -YA2 Motor nemá splněny podmínky pro opuštění pozice HOME', class Errors, trigger "DB_ALARM_OP2_M_1" bit 4
   438: 'OP2_N0 -YA2 Motor nemá splněny podmínky pro opuštění pozice WORK', class Errors, trigger "DB_ALARM_OP2_M_1" bit 5
   439: 'OP2_N0 -YA2 Motor nedojel do požadované pozice WORK', class Errors, trigger "DB_ALARM_OP2_M_1" bit 6
   440: 'OP2_N0 -YA2 Motor nedojel do požadované pozice HOME', class Errors, trigger "DB_ALARM_OP2_M_1" bit 7
   441: 'OP2_RESERVE_1 -YA2', class Errors, trigger "DB_ALARM_OP2_M_1" bit 8
   442: 'OP2_RESERVE_2 -YA2', class Errors, trigger "DB_ALARM_OP2_M_1" bit 9
   443: 'OP2_RESERVE_3 -YA2', class Errors, trigger "DB_ALARM_OP2_M_1" bit 10
   444: 'OP2_RESERVE_4 -YA2', class Errors, trigger "DB_ALARM_OP2_M_1" bit 11
   445: 'OP2_RESERVE_5 -YA2', class Errors, trigger "DB_ALARM_OP2_M_1" bit 12
   446: 'OP2_RESERVE_6 -YA2', class Errors, trigger "DB_ALARM_OP2_M_1" bit 13
   447: 'OP2_RESERVE_7 -YA2', class Errors, trigger "DB_ALARM_OP2_M_1" bit 14
   448: 'OP2_RESERVE_8 -YA2', class Errors, trigger "DB_ALARM_OP2_M_1" bit 15
   449: 'OP2_N0 -YA3 Nespecifikovaný režim motoru AUTOMAT/MANUAL', class Errors, trigger "DB_ALARM_OP2_M_2" bit 0
   450: 'OP2_N0 -YA3 Externí alarm err 1', class Errors, trigger "DB_ALARM_OP2_M_2" bit 1
   451: 'OP2_N0 -YA3 Externí alarm err 2', class Errors, trigger "DB_ALARM_OP2_M_2" bit 2
   452: 'OP2_N0 -YA3 Externí alarm err 3', class Errors, trigger "DB_ALARM_OP2_M_2" bit 3
   453: 'OP2_N0 -YA3 Motor nemá splněny podmínky pro opuštění pozice HOME', class Errors, trigger "DB_ALARM_OP2_M_2" bit 4
   454: 'OP2_N0 -YA3 Motor nemá splněny podmínky pro opuštění pozice WORK', class Errors, trigger "DB_ALARM_OP2_M_2" bit 5
   455: 'OP2_N0 -YA3 Motor nedojel do požadované pozice WORK', class Errors, trigger "DB_ALARM_OP2_M_2" bit 6
   456: 'OP2_N0 -YA3 Motor nedojel do požadované pozice HOME', class Errors, trigger "DB_ALARM_OP2_M_2" bit 7
   457: 'OP2_RESERVE_1-YA3', class Errors, trigger "DB_ALARM_OP2_M_2" bit 8
   458: 'OP2_RESERVE_2-YA3', class Errors, trigger "DB_ALARM_OP2_M_2" bit 9
   459: 'OP2_RESERVE_3-YA3', class Errors, trigger "DB_ALARM_OP2_M_2" bit 10
   460: 'OP2_RESERVE_4-YA3', class Errors, trigger "DB_ALARM_OP2_M_2" bit 11
   461: 'OP2_RESERVE_5-YA3', class Errors, trigger "DB_ALARM_OP2_M_2" bit 12
   462: 'OP2_RESERVE_6-YA3', class Errors, trigger "DB_ALARM_OP2_M_2" bit 13
   463: 'OP2_RESERVE_7-YA3', class Errors, trigger "DB_ALARM_OP2_M_2" bit 14
   464: 'OP2_RESERVE_8-YA3', class Errors, trigger "DB_ALARM_OP2_M_2" bit 15
   465: 'OP2_N0 -YA4 Nespecifikovaný režim motoru AUTOMAT/MANUAL', class Errors, trigger "DB_ALARM_OP2_M_3" bit 0
   466: 'OP2_N0 -YA4 Externí alarm err 1', class Errors, trigger "DB_ALARM_OP2_M_3" bit 1
   467: 'OP2_N0 -YA4 Externí alarm err 2', class Errors, trigger "DB_ALARM_OP2_M_3" bit 2
   468: 'OP2_N0 -YA4 Externí alarm err 3', class Errors, trigger "DB_ALARM_OP2_M_3" bit 3
   469: 'OP2_N0 -YA4 Motor nemá splněny podmínky pro opuštění pozice HOME', class Errors, trigger "DB_ALARM_OP2_M_3" bit 4
   470: 'OP2_N0 -YA4 Motor nemá splněny podmínky pro opuštění pozice WORK', class Errors, trigger "DB_ALARM_OP2_M_3" bit 5
   471: 'OP2_N0 -YA4 Motor nedojel do požadované pozice WORK', class Errors, trigger "DB_ALARM_OP2_M_3" bit 6
   472: 'OP2_N0 -YA4 Motor nedojel do požadované pozice HOME', class Errors, trigger "DB_ALARM_OP2_M_3" bit 7
   473: 'OP2_RESERVE_1-YA4', class Errors, trigger "DB_ALARM_OP2_M_3" bit 8
   474: 'OP2_RESERVE_2-YA4', class Errors, trigger "DB_ALARM_OP2_M_3" bit 9
   475: 'OP2_RESERVE_3-YA4', class Errors, trigger "DB_ALARM_OP2_M_3" bit 10
   476: 'OP2_RESERVE_4-YA4', class Errors, trigger "DB_ALARM_OP2_M_3" bit 11
   477: 'OP2_RESERVE_5-YA4', class Errors, trigger "DB_ALARM_OP2_M_3" bit 12
   478: 'OP2_RESERVE_6-YA4', class Errors, trigger "DB_ALARM_OP2_M_3" bit 13
   479: 'OP2_RESERVE_7-YA4', class Errors, trigger "DB_ALARM_OP2_M_3" bit 14
   480: 'OP2_RESERVE_8-YA4', class Errors, trigger "DB_ALARM_OP2_M_3" bit 15
   481: 'OP2_N0 -YA5 Nespecifikovaný režim motoru AUTOMAT/MANUAL', class Errors, trigger "DB_ALARM_OP2_M_4" bit 0
   482: 'OP2_N0 -YA5 Externí alarm err 1', class Errors, trigger "DB_ALARM_OP2_M_4" bit 1
   483: 'OP2_N0 -YA5 Externí alarm err 2', class Errors, trigger "DB_ALARM_OP2_M_4" bit 2
   484: 'OP2_N0 -YA5 Externí alarm err 3', class Errors, trigger "DB_ALARM_OP2_M_4" bit 3
   485: 'OP2_N0 -YA5 Motor nemá splněny podmínky pro opuštění pozice HOME', class Errors, trigger "DB_ALARM_OP2_M_4" bit 4
   486: 'OP2_N0 -YA5 Motor nemá splněny podmínky pro opuštění pozice WORK', class Errors, trigger "DB_ALARM_OP2_M_4" bit 5
   487: 'OP2_N0 -YA5 Motor nedojel do požadované pozice WORK', class Errors, trigger "DB_ALARM_OP2_M_4" bit 6
   488: 'OP2_N0 -YA5 Motor nedojel do požadované pozice HOME', class Errors, trigger "DB_ALARM_OP2_M_4" bit 7
   489: 'OP2_RESERVE_1-YA5', class Errors, trigger "DB_ALARM_OP2_M_4" bit 8
   490: 'OP2_RESERVE_2-YA5', class Errors, trigger "DB_ALARM_OP2_M_4" bit 9
   491: 'OP2_RESERVE_3-YA5', class Errors, trigger "DB_ALARM_OP2_M_4" bit 10
   492: 'OP2_RESERVE_4-YA5', class Errors, trigger "DB_ALARM_OP2_M_4" bit 11
   493: 'OP2_RESERVE_5-YA5', class Errors, trigger "DB_ALARM_OP2_M_4" bit 12
   494: 'OP2_RESERVE_6-YA5', class Errors, trigger "DB_ALARM_OP2_M_4" bit 13
   495: 'OP2_RESERVE_7-YA5', class Errors, trigger "DB_ALARM_OP2_M_4" bit 14
   496: 'OP2_RESERVE_8-YA5', class Errors, trigger "DB_ALARM_OP2_M_4" bit 15
   497: 'OP2_N0 -YA6 Nespecifikovaný režim motoru AUTOMAT/MANUAL', class Errors, trigger "DB_ALARM_OP2_M_5" bit 0
   498: 'OP2_N0 -YA6 Externí alarm err 1', class Errors, trigger "DB_ALARM_OP2_M_5" bit 1
   499: 'OP2_N0 -YA6 Externí alarm err 2', class Errors, trigger "DB_ALARM_OP2_M_5" bit 2
   500: 'OP2_N0 -YA6 Externí alarm err 3', class Errors, trigger "DB_ALARM_OP2_M_5" bit 3
   501: 'OP2_N0 -YA6 Motor nemá splněny podmínky pro opuštění pozice HOME', class Errors, trigger "DB_ALARM_OP2_M_5" bit 4
   502: 'OP2_N0 -YA6 Motor nemá splněny podmínky pro opuštění pozice WORK', class Errors, trigger "DB_ALARM_OP2_M_5" bit 5
   503: 'OP2_N0 -YA6 Motor nedojel do požadované pozice WORK', class Errors, trigger "DB_ALARM_OP2_M_5" bit 6
   504: 'OP2_N0 -YA6 Motor nedojel do požadované pozice HOME', class Errors, trigger "DB_ALARM_OP2_M_5" bit 7
   505: 'OP2_RESERVE_1-YA6', class Errors, trigger "DB_ALARM_OP2_M_5" bit 8
   506: 'OP2_RESERVE_2-YA6', class Errors, trigger "DB_ALARM_OP2_M_5" bit 9
   507: 'OP2_RESERVE_3-YA6', class Errors, trigger "DB_ALARM_OP2_M_5" bit 10
   508: 'OP2_RESERVE_4-YA6', class Errors, trigger "DB_ALARM_OP2_M_5" bit 11
   509: 'OP2_RESERVE_5-YA6', class Errors, trigger "DB_ALARM_OP2_M_5" bit 12
   510: 'OP2_RESERVE_6-YA6', class Errors, trigger "DB_ALARM_OP2_M_5" bit 13
   511: 'OP2_RESERVE_7-YA6', class Errors, trigger "DB_ALARM_OP2_M_5" bit 14
   512: 'OP2_RESERVE_8-YA6', class Errors, trigger "DB_ALARM_OP2_M_5" bit 15
   513: 'OP2_N0 -YA7 Nespecifikovaný režim motoru AUTOMAT/MANUAL', class Errors, trigger "DB_ALARM_OP2_M_6" bit 0
   514: 'OP2_N0 -YA7 Externí alarm err 1', class Errors, trigger "DB_ALARM_OP2_M_6" bit 1
   515: 'OP2_N0 -YA7 Externí alarm err 2', class Errors, trigger "DB_ALARM_OP2_M_6" bit 2
   516: 'OP2_N0 -YA7 Externí alarm err 3', class Errors, trigger "DB_ALARM_OP2_M_6" bit 3
   517: 'OP2_N0 -YA7 Motor nemá splněny podmínky pro opuštění pozice HOME', class Errors, trigger "DB_ALARM_OP2_M_6" bit 4
   518: 'OP2_N0 -YA7 Motor nemá splněny podmínky pro opuštění pozice WORK', class Errors, trigger "DB_ALARM_OP2_M_6" bit 5
   519: 'OP2_N0 -YA7 Motor nedojel do požadované pozice WORK', class Errors, trigger "DB_ALARM_OP2_M_6" bit 6
   520: 'OP2_N0 -YA7 Motor nedojel do požadované pozice HOME', class Errors, trigger "DB_ALARM_OP2_M_6" bit 7
   521: 'OP2_RESERVE_1-YA7', class Errors, trigger "DB_ALARM_OP2_M_6" bit 8
   522: 'OP2_RESERVE_2-YA7', class Errors, trigger "DB_ALARM_OP2_M_6" bit 9
   523: 'OP2_RESERVE_3-YA7', class Errors, trigger "DB_ALARM_OP2_M_6" bit 10
   524: 'OP2_RESERVE_4-YA7', class Errors, trigger "DB_ALARM_OP2_M_6" bit 11
   525: 'OP2_RESERVE_5-YA7', class Errors, trigger "DB_ALARM_OP2_M_6" bit 12
   526: 'OP2_RESERVE_6-YA7', class Errors, trigger "DB_ALARM_OP2_M_6" bit 13
   527: 'OP2_RESERVE_7-YA7', class Errors, trigger "DB_ALARM_OP2_M_6" bit 14
   528: 'OP2_RESERVE_8-YA7', class Errors, trigger "DB_ALARM_OP2_M_6" bit 15
   529: 'OP2_N0 -YA8 Nespecifikovaný režim motoru AUTOMAT/MANUAL', class Errors, trigger "DB_ALARM_OP2_M_7" bit 0
   530: 'OP2_N0 -YA8 Externí alarm err 1', class Errors, trigger "DB_ALARM_OP2_M_7" bit 1
   531: 'OP2_N0 -YA8 Externí alarm err 2', class Errors, trigger "DB_ALARM_OP2_M_7" bit 2
   532: 'OP2_N0 -YA8 Externí alarm err 3', class Errors, trigger "DB_ALARM_OP2_M_7" bit 3
   533: 'OP2_N0 -YA8 Motor nemá splněny podmínky pro opuštění pozice HOME', class Errors, trigger "DB_ALARM_OP2_M_7" bit 4
   534: 'OP2_N0 -YA8 Motor nemá splněny podmínky pro opuštění pozice WORK', class Errors, trigger "DB_ALARM_OP2_M_7" bit 5
   535: 'OP2_N0 -YA8 Motor nedojel do požadované pozice WORK', class Errors, trigger "DB_ALARM_OP2_M_7" bit 6
   536: 'OP2_N0 -YA8 Motor nedojel do požadované pozice HOME', class Errors, trigger "DB_ALARM_OP2_M_7" bit 7
   537: 'OP2_RESERVE_1-YA8', class Errors, trigger "DB_ALARM_OP2_M_7" bit 8
   538: 'OP2_RESERVE_2-YA8', class Errors, trigger "DB_ALARM_OP2_M_7" bit 9
   539: 'OP2_RESERVE_3-YA8', class Errors, trigger "DB_ALARM_OP2_M_7" bit 10
   540: 'OP2_RESERVE_4-YA8', class Errors, trigger "DB_ALARM_OP2_M_7" bit 11
   541: 'OP2_RESERVE_5-YA8', class Errors, trigger "DB_ALARM_OP2_M_7" bit 12
   542: 'OP2_RESERVE_6-YA8', class Errors, trigger "DB_ALARM_OP2_M_7" bit 13
   543: 'OP2_RESERVE_7-YA8', class Errors, trigger "DB_ALARM_OP2_M_7" bit 14
   544: 'OP2_RESERVE_8-YA8', class Errors, trigger "DB_ALARM_OP2_M_7" bit 15
   545: 'OP2_N0 Nespecifikovaný režim motoru AUTOMAT/MANUAL', class Errors, trigger "DB_ALARM_OP2_M_8" bit 0
   546: 'OP2_N0 Externí alarm err 1', class Errors, trigger "DB_ALARM_OP2_M_8" bit 1
   547: 'OP2_N0 Externí alarm err 2', class Errors, trigger "DB_ALARM_OP2_M_8" bit 2
   548: 'OP2_N0 Externí alarm err 3', class Errors, trigger "DB_ALARM_OP2_M_8" bit 3
   549: 'OP2_N0 Motor nemá splněny podmínky pro opuštění pozice HOME', class Errors, trigger "DB_ALARM_OP2_M_8" bit 4
   550: 'OP2_N0 Motor nemá splněny podmínky pro opuštění pozice WORK', class Errors, trigger "DB_ALARM_OP2_M_8" bit 5
   551: 'OP2_N0 Motor nedojel do požadované pozice WORK', class Errors, trigger "DB_ALARM_OP2_M_8" bit 6
   552: 'OP2_N0 Motor nedojel do požadované pozice HOME', class Errors, trigger "DB_ALARM_OP2_M_8" bit 7
   553: 'OP2_RESERVE_1', class Errors, trigger "DB_ALARM_OP2_M_8" bit 8
   554: 'OP2_RESERVE_2', class Errors, trigger "DB_ALARM_OP2_M_8" bit 9
   555: 'OP2_RESERVE_3', class Errors, trigger "DB_ALARM_OP2_M_8" bit 10
   556: 'OP2_RESERVE_4', class Errors, trigger "DB_ALARM_OP2_M_8" bit 11
   557: 'OP2_RESERVE_5', class Errors, trigger "DB_ALARM_OP2_M_8" bit 12
   558: 'OP2_RESERVE_6', class Errors, trigger "DB_ALARM_OP2_M_8" bit 13
   559: 'OP2_RESERVE_7', class Errors, trigger "DB_ALARM_OP2_M_8" bit 14
   560: 'OP2_RESERVE_8', class Errors, trigger "DB_ALARM_OP2_M_8" bit 15
   561: 'OP2_N0 Nespecifikovaný režim motoru AUTOMAT/MANUAL', class Errors, trigger "DB_ALARM_OP2_M_9" bit 0
   562: 'OP2_N0 Externí alarm err 1', class Errors, trigger "DB_ALARM_OP2_M_9" bit 1
   563: 'OP2_N0 Externí alarm err 2', class Errors, trigger "DB_ALARM_OP2_M_9" bit 2
   564: 'OP2_N0 Externí alarm err 3', class Errors, trigger "DB_ALARM_OP2_M_9" bit 3
   565: 'OP2_N0 Motor nemá splněny podmínky pro opuštění pozice HOME', class Errors, trigger "DB_ALARM_OP2_M_9" bit 4
   566: 'OP2_N0 Motor nemá splněny podmínky pro opuštění pozice WORK', class Errors, trigger "DB_ALARM_OP2_M_9" bit 5
   567: 'OP2_N0 Motor nedojel do požadované pozice WORK', class Errors, trigger "DB_ALARM_OP2_M_9" bit 6
   568: 'OP2_N0 Motor nedojel do požadované pozice HOME', class Errors, trigger "DB_ALARM_OP2_M_9" bit 7
   569: 'OP2_RESERVE_1', class Errors, trigger "DB_ALARM_OP2_M_9" bit 8
   570: 'OP2_RESERVE_2', class Errors, trigger "DB_ALARM_OP2_M_9" bit 9
   571: 'OP2_RESERVE_3', class Errors, trigger "DB_ALARM_OP2_M_9" bit 10
   572: 'OP2_RESERVE_4', class Errors, trigger "DB_ALARM_OP2_M_9" bit 11
   573: 'OP2_RESERVE_5', class Errors, trigger "DB_ALARM_OP2_M_9" bit 12
   574: 'OP2_RESERVE_6', class Errors, trigger "DB_ALARM_OP2_M_9" bit 13
   575: 'OP2_RESERVE_7', class Errors, trigger "DB_ALARM_OP2_M_9" bit 14
   576: 'OP2_RESERVE_8', class Errors, trigger "DB_ALARM_OP2_M_9" bit 15
   577: 'OP2_N0 Nespecifikovaný režim motoru AUTOMAT/MANUAL', class Errors, trigger "DB_ALARM_OP2_M_10" bit 0
   578: 'OP2_N0 Externí alarm err 1', class Errors, trigger "DB_ALARM_OP2_M_10" bit 1
   579: 'OP2_N0 Externí alarm err 2', class Errors, trigger "DB_ALARM_OP2_M_10" bit 2
   580: 'OP2_N0 Externí alarm err 3', class Errors, trigger "DB_ALARM_OP2_M_10" bit 3
   581: 'OP2_N0 Motor nemá splněny podmínky pro opuštění pozice HOME', class Errors, trigger "DB_ALARM_OP2_M_10" bit 4
   582: 'OP2_N0 Motor nemá splněny podmínky pro opuštění pozice WORK', class Errors, trigger "DB_ALARM_OP2_M_10" bit 5
   583: 'OP2_N0 Motor nedojel do požadované pozice WORK', class Errors, trigger "DB_ALARM_OP2_M_10" bit 6
   584: 'OP2_N0 Motor nedojel do požadované pozice HOME', class Errors, trigger "DB_ALARM_OP2_M_10" bit 7
   585: 'OP2_RESERVE_1', class Errors, trigger "DB_ALARM_OP2_M_10" bit 8
   586: 'OP2_RESERVE_2', class Errors, trigger "DB_ALARM_OP2_M_10" bit 9
   587: 'OP2_RESERVE_3', class Errors, trigger "DB_ALARM_OP2_M_10" bit 10
   588: 'OP2_RESERVE_4', class Errors, trigger "DB_ALARM_OP2_M_10" bit 11
   589: 'OP2_RESERVE_5', class Errors, trigger "DB_ALARM_OP2_M_10" bit 12
   590: 'OP2_RESERVE_6', class Errors, trigger "DB_ALARM_OP2_M_10" bit 13
   591: 'OP2_RESERVE_7', class Errors, trigger "DB_ALARM_OP2_M_10" bit 14
   592: 'OP2_RESERVE_8', class Errors, trigger "DB_ALARM_OP2_M_10" bit 15
   593: 'OP2_N0 Nespecifikovaný režim motoru AUTOMAT/MANUAL', class Errors, trigger "DB_ALARM_OP2_M_11" bit 0
   594: 'OP2_N0 Externí alarm err 1', class Errors, trigger "DB_ALARM_OP2_M_11" bit 1
   595: 'OP2_N0 Externí alarm err 2', class Errors, trigger "DB_ALARM_OP2_M_11" bit 2
   596: 'OP2_N0 Externí alarm err 3', class Errors, trigger "DB_ALARM_OP2_M_11" bit 3
   597: 'OP2_N0 Motor nemá splněny podmínky pro opuštění pozice HOME', class Errors, trigger "DB_ALARM_OP2_M_11" bit 4
   598: 'OP2_N0 Motor nemá splněny podmínky pro opuštění pozice WORK', class Errors, trigger "DB_ALARM_OP2_M_11" bit 5
   599: 'OP2_N0 Motor nedojel do požadované pozice WORK', class Errors, trigger "DB_ALARM_OP2_M_11" bit 6
   600: 'OP2_N0 Motor nedojel do požadované pozice HOME', class Errors, trigger "DB_ALARM_OP2_M_11" bit 7
   601: 'OP2_RESERVE_1', class Errors, trigger "DB_ALARM_OP2_M_11" bit 8
   602: 'OP2_RESERVE_2', class Errors, trigger "DB_ALARM_OP2_M_11" bit 9
   603: 'OP2_RESERVE_3', class Errors, trigger "DB_ALARM_OP2_M_11" bit 10
   604: 'OP2_RESERVE_4', class Errors, trigger "DB_ALARM_OP2_M_11" bit 11
   605: 'OP2_RESERVE_5', class Errors, trigger "DB_ALARM_OP2_M_11" bit 12
   606: 'OP2_RESERVE_6', class Errors, trigger "DB_ALARM_OP2_M_11" bit 13
   607: 'OP2_RESERVE_7', class Errors, trigger "DB_ALARM_OP2_M_11" bit 14
   608: 'OP2_RESERVE_8', class Errors, trigger "DB_ALARM_OP2_M_11" bit 15
   609: 'OP2_N0 Nespecifikovaný režim motoru AUTOMAT/MANUAL', class Errors, trigger "DB_ALARM_OP2_M_12" bit 0
   610: 'OP2_N0 Externí alarm err 1', class Errors, trigger "DB_ALARM_OP2_M_12" bit 1
   611: 'OP2_N0 Externí alarm err 2', class Errors, trigger "DB_ALARM_OP2_M_12" bit 2
   612: 'OP2_N0 Externí alarm err 3', class Errors, trigger "DB_ALARM_OP2_M_12" bit 3
   613: 'OP2_N0 Motor nemá splněny podmínky pro opuštění pozice HOME', class Errors, trigger "DB_ALARM_OP2_M_12" bit 4
   614: 'OP2_N0 Motor nemá splněny podmínky pro opuštění pozice WORK', class Errors, trigger "DB_ALARM_OP2_M_12" bit 5
   615: 'OP2_N0 Motor nedojel do požadované pozice WORK', class Errors, trigger "DB_ALARM_OP2_M_12" bit 6
   616: 'OP2_N0 Motor nedojel do požadované pozice HOME', class Errors, trigger "DB_ALARM_OP2_M_12" bit 7
   617: 'OP2_RESERVE_1', class Errors, trigger "DB_ALARM_OP2_M_12" bit 8
   618: 'OP2_RESERVE_2', class Errors, trigger "DB_ALARM_OP2_M_12" bit 9
   619: 'OP2_RESERVE_3', class Errors, trigger "DB_ALARM_OP2_M_12" bit 10
   620: 'OP2_RESERVE_4', class Errors, trigger "DB_ALARM_OP2_M_12" bit 11
   621: 'OP2_RESERVE_5', class Errors, trigger "DB_ALARM_OP2_M_12" bit 12
   622: 'OP2_RESERVE_6', class Errors, trigger "DB_ALARM_OP2_M_12" bit 13
   623: 'OP2_RESERVE_7', class Errors, trigger "DB_ALARM_OP2_M_12" bit 14
   624: 'OP2_RESERVE_8', class Errors, trigger "DB_ALARM_OP2_M_12" bit 15
   625: 'OP2_N0 Nespecifikovaný režim motoru AUTOMAT/MANUAL', class Errors, trigger "DB_ALARM_OP2_M_13" bit 0
   626: 'OP2_N0 Externí alarm err 1', class Errors, trigger "DB_ALARM_OP2_M_13" bit 1
   627: 'OP2_N0 Externí alarm err 2', class Errors, trigger "DB_ALARM_OP2_M_13" bit 2
   628: 'OP2_N0 Externí alarm err 3', class Errors, trigger "DB_ALARM_OP2_M_13" bit 3
   629: 'OP2_N0 Motor nemá splněny podmínky pro opuštění pozice HOME', class Errors, trigger "DB_ALARM_OP2_M_13" bit 4
   630: 'OP2_N0 Motor nemá splněny podmínky pro opuštění pozice WORK', class Errors, trigger "DB_ALARM_OP2_M_13" bit 5
   631: 'OP2_N0 Motor nedojel do požadované pozice WORK', class Errors, trigger "DB_ALARM_OP2_M_13" bit 6
   632: 'OP2_N0 Motor nedojel do požadované pozice HOME', class Errors, trigger "DB_ALARM_OP2_M_13" bit 7
   633: 'OP2_RESERVE_1', class Errors, trigger "DB_ALARM_OP2_M_13" bit 8
   634: 'OP2_RESERVE_2', class Errors, trigger "DB_ALARM_OP2_M_13" bit 9
   635: 'OP2_RESERVE_3', class Errors, trigger "DB_ALARM_OP2_M_13" bit 10
   636: 'OP2_RESERVE_4', class Errors, trigger "DB_ALARM_OP2_M_13" bit 11
   637: 'OP2_RESERVE_5', class Errors, trigger "DB_ALARM_OP2_M_13" bit 12
   638: 'OP2_RESERVE_6', class Errors, trigger "DB_ALARM_OP2_M_13" bit 13
   639: 'OP2_RESERVE_7', class Errors, trigger "DB_ALARM_OP2_M_13" bit 14
   640: 'OP2_RESERVE_8', class Errors, trigger "DB_ALARM_OP2_M_13" bit 15
   641: 'OP2_N0 Nespecifikovaný režim motoru AUTOMAT/MANUAL', class Errors, trigger "DB_ALARM_OP2_M_14" bit 0
   642: 'OP2_N0 Externí alarm err 1', class Errors, trigger "DB_ALARM_OP2_M_14" bit 1
   643: 'OP2_N0 Externí alarm err 2', class Errors, trigger "DB_ALARM_OP2_M_14" bit 2
   644: 'OP2_N0 Externí alarm err 3', class Errors, trigger "DB_ALARM_OP2_M_14" bit 3
   645: 'OP2_N0 Motor nemá splněny podmínky pro opuštění pozice HOME', class Errors, trigger "DB_ALARM_OP2_M_14" bit 4
   646: 'OP2_N0 Motor nemá splněny podmínky pro opuštění pozice WORK', class Errors, trigger "DB_ALARM_OP2_M_14" bit 5
   647: 'OP2_N0 Motor nedojel do požadované pozice WORK', class Errors, trigger "DB_ALARM_OP2_M_14" bit 6
   648: 'OP2_N0 Motor nedojel do požadované pozice HOME', class Errors, trigger "DB_ALARM_OP2_M_14" bit 7
   649: 'OP2_RESERVE_1', class Errors, trigger "DB_ALARM_OP2_M_14" bit 8
   650: 'OP2_RESERVE_2', class Errors, trigger "DB_ALARM_OP2_M_14" bit 9
   651: 'OP2_RESERVE_3', class Errors, trigger "DB_ALARM_OP2_M_14" bit 10
   652: 'OP2_RESERVE_4', class Errors, trigger "DB_ALARM_OP2_M_14" bit 11
   653: 'OP2_RESERVE_5', class Errors, trigger "DB_ALARM_OP2_M_14" bit 12
   654: 'OP2_RESERVE_6', class Errors, trigger "DB_ALARM_OP2_M_14" bit 13
   655: 'OP2_RESERVE_7', class Errors, trigger "DB_ALARM_OP2_M_14" bit 14
   656: 'OP2_RESERVE_8', class Errors, trigger "DB_ALARM_OP2_M_14" bit 15
   657: 'OP2_N0 Nespecifikovaný režim motoru AUTOMAT/MANUAL', class Errors, trigger "DB_ALARM_OP2_M_15" bit 0
   658: 'OP2_N0 Externí alarm err 1', class Errors, trigger "DB_ALARM_OP2_M_15" bit 1
   659: 'OP2_N0 Externí alarm err 2', class Errors, trigger "DB_ALARM_OP2_M_15" bit 2
   660: 'OP2_N0 Externí alarm err 3', class Errors, trigger "DB_ALARM_OP2_M_15" bit 3
   661: 'OP2_N0 Motor nemá splněny podmínky pro opuštění pozice HOME', class Errors, trigger "DB_ALARM_OP2_M_15" bit 4
   662: 'OP2_N0 Motor nemá splněny podmínky pro opuštění pozice WORK', class Errors, trigger "DB_ALARM_OP2_M_15" bit 5
   663: 'OP2_N0 Motor nedojel do požadované pozice WORK', class Errors, trigger "DB_ALARM_OP2_M_15" bit 6
   664: 'OP2_N0 Motor nedojel do požadované pozice HOME', class Errors, trigger "DB_ALARM_OP2_M_15" bit 7
   665: 'OP2_RESERVE_1', class Errors, trigger "DB_ALARM_OP2_M_15" bit 8
   666: 'OP2_RESERVE_2', class Errors, trigger "DB_ALARM_OP2_M_15" bit 9
   667: 'OP2_RESERVE_3', class Errors, trigger "DB_ALARM_OP2_M_15" bit 10
   668: 'OP2_RESERVE_4', class Errors, trigger "DB_ALARM_OP2_M_15" bit 11
   669: 'OP2_RESERVE_5', class Errors, trigger "DB_ALARM_OP2_M_15" bit 12
   670: 'OP2_RESERVE_6', class Errors, trigger "DB_ALARM_OP2_M_15" bit 13
   671: 'OP2_RESERVE_7', class Errors, trigger "DB_ALARM_OP2_M_15" bit 14
   672: 'OP2_RESERVE_8', class Errors, trigger "DB_ALARM_OP2_M_15" bit 15
   673: 'OP3_N0 -YB1 Nespecifikovaný režim motoru AUTOMAT/MANUAL', class Errors, trigger "DB_ALARM_OP3_M_0" bit 0
   674: 'OP3_N0 -YB1 Externí alarm err 1', class Errors, trigger "DB_ALARM_OP3_M_0" bit 1
   675: 'OP3_N0 -YB1 Externí alarm err 2', class Errors, trigger "DB_ALARM_OP3_M_0" bit 2
   676: 'OP3_N0 -YB1 Externí alarm err 3', class Errors, trigger "DB_ALARM_OP3_M_0" bit 3
   677: 'OP3_N0 -YB1 Motor nemá splněny podmínky pro opuštění pozice HOME', class Errors, trigger "DB_ALARM_OP3_M_0" bit 4
   678: 'OP3_N0 -YB1 Motor nemá splněny podmínky pro opuštění pozice WORK', class Errors, trigger "DB_ALARM_OP3_M_0" bit 5
   679: 'OP3_N0 -YB1 Motor nedojel do požadované pozice WORK', class Errors, trigger "DB_ALARM_OP3_M_0" bit 6
   680: 'OP3_N0 -YB1 Motor nedojel do požadované pozice HOME', class Errors, trigger "DB_ALARM_OP3_M_0" bit 7
   681: '-YB1 OP3_RESERVE_1', class Errors, trigger "DB_ALARM_OP3_M_0" bit 8
   682: '-YB1 OP3_RESERVE_2', class Errors, trigger "DB_ALARM_OP3_M_0" bit 9
   683: '-YB1 OP3_RESERVE_3', class Errors, trigger "DB_ALARM_OP3_M_0" bit 10
   684: '-YB1 OP3_RESERVE_4', class Errors, trigger "DB_ALARM_OP3_M_0" bit 11
   685: '-YB1 OP3_RESERVE_5', class Errors, trigger "DB_ALARM_OP3_M_0" bit 12
   686: '-YB1 OP3_RESERVE_6', class Errors, trigger "DB_ALARM_OP3_M_0" bit 13
   687: '-YB1 OP3_RESERVE_7', class Errors, trigger "DB_ALARM_OP3_M_0" bit 14
   688: '-YB1 OP3_RESERVE_8', class Errors, trigger "DB_ALARM_OP3_M_0" bit 15
   689: 'OP3_N0 -YB2 Nespecifikovaný režim motoru AUTOMAT/MANUAL', class Errors, trigger "DB_ALARM_OP3_M_1" bit 0
   690: 'OP3_N0 -YB2 Externí alarm err 1', class Errors, trigger "DB_ALARM_OP3_M_1" bit 1
   691: 'OP3_N0 -YB2 Externí alarm err 2', class Errors, trigger "DB_ALARM_OP3_M_1" bit 2
   692: 'OP3_N0 -YB2 Externí alarm err 3', class Errors, trigger "DB_ALARM_OP3_M_1" bit 3
   693: 'OP3_N0 -YB2 Motor nemá splněny podmínky pro opuštění pozice HOME', class Errors, trigger "DB_ALARM_OP3_M_1" bit 4
   694: 'OP3_N0 -YB2 Motor nemá splněny podmínky pro opuštění pozice WORK', class Errors, trigger "DB_ALARM_OP3_M_1" bit 5
   695: 'OP3_N0 -YB2 Motor nedojel do požadované pozice WORK', class Errors, trigger "DB_ALARM_OP3_M_1" bit 6
   696: 'OP3_N0 -YB2 Motor nedojel do požadované pozice HOME', class Errors, trigger "DB_ALARM_OP3_M_1" bit 7
   697: '-YB2 OP3_RESERVE_1', class Errors, trigger "DB_ALARM_OP3_M_1" bit 8
   698: '-YB2 OP3_RESERVE_2', class Errors, trigger "DB_ALARM_OP3_M_1" bit 9
   699: '-YB2 OP3_RESERVE_3', class Errors, trigger "DB_ALARM_OP3_M_1" bit 10
   700: '-YB2 OP3_RESERVE_4', class Errors, trigger "DB_ALARM_OP3_M_1" bit 11
   701: '-YB2 OP3_RESERVE_5', class Errors, trigger "DB_ALARM_OP3_M_1" bit 12
   702: '-YB2 OP3_RESERVE_6', class Errors, trigger "DB_ALARM_OP3_M_1" bit 13
   703: '-YB2 OP3_RESERVE_7', class Errors, trigger "DB_ALARM_OP3_M_1" bit 14
   704: '-YB2 OP3_RESERVE_8', class Errors, trigger "DB_ALARM_OP3_M_1" bit 15
   705: 'OP3_N0 -YB3 Nespecifikovaný režim motoru AUTOMAT/MANUAL', class Errors, trigger "DB_ALARM_OP3_M_2" bit 0
   706: 'OP3_N0 -YB3 Externí alarm err 1', class Errors, trigger "DB_ALARM_OP3_M_2" bit 1
   707: 'OP3_N0 -YB3 Externí alarm err 2', class Errors, trigger "DB_ALARM_OP3_M_2" bit 2
   708: 'OP3_N0 -YB3 Externí alarm err 3', class Errors, trigger "DB_ALARM_OP3_M_2" bit 3
   709: 'OP3_N0 -YB3 Motor nemá splněny podmínky pro opuštění pozice HOME', class Errors, trigger "DB_ALARM_OP3_M_2" bit 4
   710: 'OP3_N0 -YB3 Motor nemá splněny podmínky pro opuštění pozice WORK', class Errors, trigger "DB_ALARM_OP3_M_2" bit 5
   711: 'OP3_N0 -YB3 Motor nedojel do požadované pozice WORK', class Errors, trigger "DB_ALARM_OP3_M_2" bit 6
   712: 'OP3_N0 -YB3 Motor nedojel do požadované pozice HOME', class Errors, trigger "DB_ALARM_OP3_M_2" bit 7
   713: '-YB3 OP3_RESERVE_1', class Errors, trigger "DB_ALARM_OP3_M_2" bit 8
   714: '-YB3 OP3_RESERVE_2', class Errors, trigger "DB_ALARM_OP3_M_2" bit 9
   715: '-YB3 OP3_RESERVE_3', class Errors, trigger "DB_ALARM_OP3_M_2" bit 10
   716: '-YB3 OP3_RESERVE_4', class Errors, trigger "DB_ALARM_OP3_M_2" bit 11
   717: '-YB3 OP3_RESERVE_5', class Errors, trigger "DB_ALARM_OP3_M_2" bit 12
   718: '-YB3 OP3_RESERVE_6', class Errors, trigger "DB_ALARM_OP3_M_2" bit 13
   719: '-YB3 OP3_RESERVE_7', class Errors, trigger "DB_ALARM_OP3_M_2" bit 14
   720: '-YB3 OP3_RESERVE_8', class Errors, trigger "DB_ALARM_OP3_M_2" bit 15
   721: 'OP3_N0 -YB4 Nespecifikovaný režim motoru AUTOMAT/MANUAL', class Errors, trigger "DB_ALARM_OP3_M_3" bit 0
   722: 'OP3_N0 -YB4 Externí alarm err 1', class Errors, trigger "DB_ALARM_OP3_M_3" bit 1
   723: 'OP3_N0 -YB4 Externí alarm err 2', class Errors, trigger "DB_ALARM_OP3_M_3" bit 2
   724: 'OP3_N0 -YB4 Externí alarm err 3', class Errors, trigger "DB_ALARM_OP3_M_3" bit 3
   725: 'OP3_N0 -YB4 Motor nemá splněny podmínky pro opuštění pozice HOME', class Errors, trigger "DB_ALARM_OP3_M_3" bit 4
   726: 'OP3_N0 -YB4 Motor nemá splněny podmínky pro opuštění pozice WORK', class Errors, trigger "DB_ALARM_OP3_M_3" bit 5
   727: 'OP3_N0 -YB4 Motor nedojel do požadované pozice WORK', class Errors, trigger "DB_ALARM_OP3_M_3" bit 6
   728: 'OP3_N0 -YB4 Motor nedojel do požadované pozice HOME', class Errors, trigger "DB_ALARM_OP3_M_3" bit 7
